(* IEC 61131-3 sources: daoli-st-library/DL_MathData (part 4) *)

(* ---- FC_DL_OrificeFlowCalc.st ---- *)
(*==============================================================================
 * 组件名称 (Component)  : FC_DL_OrificeFlowCalc
 * 所属子库 (Sublibrary) : DL_MathData
 * 当前版本 (Version)    : 1.0.0
 * 兼容性 (Platform)     : CODESYS 3.5 / TwinCAT 3 / 汇川 InoProShop / Machine Expert
 *                         仅依赖纯 IEC 61131-3 标准元素，零厂商方言
 * 功能描述 (Function)   : 孔板差压流量计算：温压补偿 + 开方 + 量程归一。
 *                         fFlow = fKCoefficient * sqrt( dP * rho(T,P) )，
 *                         密度委托 FC_DL_AirDensity（理想气体同源式，RH=0 干气口径），
 *                         开方委托 FC_DL_NthRoot(2)，本函数只做前置校验 + 钳位 + 错误码，
 *                         不重写任何开方/密度数学内核（T0 红线）。
 * 溯源 (Origin)         : 道莅 clean-room 防御性实现
 * 本文件内含 (Contains) : TYPE E_DL_MathErr / FUNCTION FC_DL_OrificeFlowCalc
 * 依赖 (Depends)        : DL_Algo/FC_DL_AirDensity、DL_MathData/FC_DL_NthRoot
 * 红线自检 (Redline)    : 无外部全局变量、无硬件地址直引 ｜ 全变量中英双语同行注释
 *                         防除零 + 量程钳位 + 非有限值防御 ｜ 枚举成员全部显式赋值
 *                         纯函数无状态保持 ｜ 输出在每条早退路径前已赋确定值
 * 错误码表 (Codes)      : 16#0001_0471 故障级 输入无效(NaN/Inf 或系数/量程非法)
 *                         16#0001_0472 故障级 差压为负
 *                         16#0001_0473 信息级 温度越界(已钳制)
 *                         16#0001_0474 信息级 压力越界(已钳制)
 *                         16#0001_0475 成功
 * 修订历史 (Revision)   : 2026-11-17  v1.0.0  首版入库 · R27 · 阶段三批 1
 * 验收向量 (Acceptance) : dP=25000 Pa, P=101325 Pa, T=20 C, K=1.0 → rho≈1.2041,
 *                         flow≈sqrt(25000*1.2041)≈173.38 m3/h，返回 0475
 *============================================================================*)

(*-----------------------------------------------------------------------------
 * 枚举: E_DL_MathErr（归属 DL_MathData，与 FC_DL_OrificeFlowCalc 同文件）
 *----------------------------------------------------------------------------*)
TYPE E_DL_MathErr :
(
    eInvalidInput := 16#0001_0471,   // 故障级：输入无效（非有限值或系数非法）/ Fault: invalid input
    eDiffPressNeg := 16#0001_0472,   // 故障级：差压为负，物理不可实现 / Fault: negative differential pressure
    eTempClamped  := 16#0001_0473,   // 信息级：温度越界已钳制 / Info: temperature clamped
    ePressClamped := 16#0001_0474,   // 信息级：压力越界已钳制 / Info: pressure clamped
    eOk           := 16#0001_0475    // 成功 / Success
);
END_TYPE

(*==============================================================================
 * 函数: FC_DL_OrificeFlowCalc（纯函数，无任何状态保持）
 * 调用约定: 每周期按需调用；返回值 = 计算有效标志。
 *============================================================================*)
FUNCTION FC_DL_OrificeFlowCalc : BOOL
VAR_INPUT
    fDiffPress_Pa  : REAL;              // 差压 [Pa]，有效域 0~50000 / Differential pressure [Pa]
    fAbsPress_Pa   : REAL;              // 绝压 [Pa]，有效域 5.0E4~2.0E6 / Absolute pressure [Pa]
    fTemp_C        : REAL;              // 温度 [摄氏度]，有效域 -40~400 / Temperature [degC]
    fKCoefficient  : REAL;              // 流量系数（含流出系数 C 的合成值），须 > 0 / Flow coefficient including discharge factor, must be > 0
    fFlowRangeMax  : REAL;              // 流量满量程 [立方米每小时]，须 > 0 / Full-scale flow [m3/h], must be > 0
END_VAR
VAR_OUTPUT
    fFlow_m3h      : REAL;              // 体积流量 [立方米每小时] / Volume flow [m3/h]
    eError         : E_DL_MathErr;      // 错误码 / Error code
END_VAR
VAR CONSTANT
    DL_ORIF_DP_MAX    : REAL := 50000.0;   // 差压量程上限 [帕] / Differential pressure span limit [Pa]
    DL_ORIF_T_MIN     : REAL := -40.0;     // 温度域下限 [摄氏度] / Temperature domain lower bound [degC]
    DL_ORIF_T_MAX     : REAL := 400.0;     // 温度域上限 [摄氏度] / Temperature domain upper bound [degC]
    DL_ORIF_P_MIN     : REAL := 5.0E4;     // 绝压域下限 [帕] / Absolute pressure lower bound [Pa]
    DL_ORIF_P_MAX     : REAL := 2.0E6;     // 绝压域上限 [帕] / Absolute pressure upper bound [Pa]
    DL_ORIF_RH_DRY    : REAL := 0.0;       // 干气口径相对湿度（委托密度入口）[%] / Dry-gas humidity fed to the density delegate [%]
    DL_ORIF_INF_MAX   : REAL := 1.0E30;    // 非有限值判定幅值上限 / Magnitude bound for finite-value check
    DL_ORIF_ZERO      : REAL := 0.0;       // 零值常量，避免裸字面量 / Zero constant, avoids a bare literal
    DL_ORIF_RHO_MIN   : LREAL := 1.0E-9;   // 密度可信下限 [千克每立方米] / Density trust lower bound [kg/m3]
END_VAR
VAR
    fDpUse    : REAL;                    // 生效差压（校验后）[帕] / Effective differential pressure [Pa]
    fTempUse  : REAL;                    // 生效温度（钳位后）[摄氏度] / Effective temperature [degC]
    fPressUse : REAL;                    // 生效绝压（钳位后）[帕] / Effective absolute pressure [Pa]
    fRho      : LREAL;                   // 委托密度输出 [千克每立方米] / Density from the delegate [kg/m3]
    fRadicand : LREAL;                   // 开方被开方数 [帕·千克每立方米] / Radicand [Pa*kg/m3]
    fRootVal  : LREAL;                   // 委托开方输出 [无量纲合成] / Square root from the delegate
    bRootOk   : BOOL;                    // 委托开方有效标志 / Delegate root validity flag
    bNonFin   : BOOL;                    // 非有限输入汇总标志 / Non-finite input aggregate flag
END_VAR

(*------------------------------------------------------------------------------
 * 段 1｜出口默认值：任何早退路径前输出已确定（哨兵 0 流量 + 输入无效码）
 *----------------------------------------------------------------------------*)
FC_DL_OrificeFlowCalc := FALSE;                       // 返回值默认无效 / return defaults to invalid
fFlow_m3h := DL_ORIF_ZERO;                            // 流量哨兵 0 / flow sentinel zero
eError := E_DL_MathErr.eInvalidInput;                 // 默认输入无效码 / default invalid-input code

(*------------------------------------------------------------------------------
 * 段 2｜非有限值闸：NaN 用自反判（x <> x），溢出用幅值上限判
 *----------------------------------------------------------------------------*)
bNonFin := (fDiffPress_Pa <> fDiffPress_Pa) OR (ABS(fDiffPress_Pa) > DL_ORIF_INF_MAX)
        OR (fAbsPress_Pa  <> fAbsPress_Pa)  OR (ABS(fAbsPress_Pa)  > DL_ORIF_INF_MAX)
        OR (fTemp_C       <> fTemp_C)       OR (ABS(fTemp_C)       > DL_ORIF_INF_MAX)
        OR (fKCoefficient <> fKCoefficient) OR (ABS(fKCoefficient) > DL_ORIF_INF_MAX)
        OR (fFlowRangeMax <> fFlowRangeMax) OR (ABS(fFlowRangeMax) > DL_ORIF_INF_MAX);
IF bNonFin THEN
    RETURN;                                           // 早退：保持默认输出 / early exit with defaults
END_IF

(*------------------------------------------------------------------------------
 * 段 3｜配置与符号闸：系数/量程必须为正，差压不允许为负
 *----------------------------------------------------------------------------*)
IF (fKCoefficient <= DL_ORIF_ZERO) OR (fFlowRangeMax <= DL_ORIF_ZERO) THEN
    RETURN;                                           // 配置非法：保持输入无效码 / invalid configuration
END_IF
IF fDiffPress_Pa < DL_ORIF_ZERO THEN
    eError := E_DL_MathErr.eDiffPressNeg;             // 故障级：差压为负 / fault: negative dp
    RETURN;
END_IF
fDpUse := fDiffPress_Pa;                              // 差压非负直接采用 / non-negative dp adopted

(*------------------------------------------------------------------------------
 * 段 4｜温度/压力钳位（信息级越界码，先到先得但压力优先级低：温度先判）
 *----------------------------------------------------------------------------*)
eError := E_DL_MathErr.eOk;                           // 预置成功 / preset success
fTempUse := fTemp_C;                                  // 温度工作副本 / temperature working copy
IF fTempUse < DL_ORIF_T_MIN THEN
    fTempUse := DL_ORIF_T_MIN;                        // 下限钳位 / floored
    eError := E_DL_MathErr.eTempClamped;              // 信息级：温度越界 / info: temperature clamped
ELSIF fTempUse > DL_ORIF_T_MAX THEN
    fTempUse := DL_ORIF_T_MAX;                        // 上限钳位 / capped
    eError := E_DL_MathErr.eTempClamped;              // 信息级：温度越界 / info: temperature clamped
END_IF
fPressUse := fAbsPress_Pa;                            // 压力工作副本 / pressure working copy
IF fPressUse < DL_ORIF_P_MIN THEN
    fPressUse := DL_ORIF_P_MIN;                       // 下限钳位 / floored
    IF eError = E_DL_MathErr.eOk THEN
        eError := E_DL_MathErr.ePressClamped;         // 信息级：压力越界（不覆盖温度码）/ info: pressure clamped
    END_IF
ELSIF fPressUse > DL_ORIF_P_MAX THEN
    fPressUse := DL_ORIF_P_MAX;                       // 上限钳位 / capped
    IF eError = E_DL_MathErr.eOk THEN
        eError := E_DL_MathErr.ePressClamped;         // 信息级：压力越界（不覆盖温度码）/ info: pressure clamped
    END_IF
END_IF

(*------------------------------------------------------------------------------
 * 段 5｜委托密度（理想气体同源式，RH=0 干气口径；委托 FC_DL_AirDensity）
 *----------------------------------------------------------------------------*)
fRho := FC_DL_AirDensity(fTempC := REAL_TO_LREAL(fTempUse), fPressPa := REAL_TO_LREAL(fPressUse), fRh := REAL_TO_LREAL(DL_ORIF_RH_DRY));   // 密度委托 [千克每立方米] / density via delegate
IF (fRho <> fRho) OR (ABS(fRho) > REAL_TO_LREAL(DL_ORIF_INF_MAX)) OR (fRho <= DL_ORIF_RHO_MIN) THEN
    eError := E_DL_MathErr.eInvalidInput;             // 委托输出不可信：按输入无效处置 / unusable delegate output
    fFlow_m3h := DL_ORIF_ZERO;                        // 流量哨兵 / flow sentinel
    FC_DL_OrificeFlowCalc := FALSE;                   // 返回无效 / return invalid
    RETURN;
END_IF

(*------------------------------------------------------------------------------
 * 段 6｜委托开方（FC_DL_NthRoot(2)）：被开方数 = 差压 x 密度，段 5 已保证非负
 *----------------------------------------------------------------------------*)
fRadicand := REAL_TO_LREAL(fDpUse) * fRho;                     // 被开方数 [帕·千克每立方米] / radicand
fRootVal := FC_DL_NthRoot(fValue := fRadicand, nRoot := 2, bValid => bRootOk);   // 开方委托 / root via delegate
IF (NOT bRootOk) OR (fRootVal <> fRootVal) OR (ABS(fRootVal) > REAL_TO_LREAL(DL_ORIF_INF_MAX)) THEN
    eError := E_DL_MathErr.eInvalidInput;             // 委托失败按输入无效处置 / delegate failure mapped to invalid input
    FC_DL_OrificeFlowCalc := FALSE;                   // 返回无效 / return invalid
    RETURN;
END_IF

(*------------------------------------------------------------------------------
 * 段 7｜量程换算与上限钳制：flow = K x root，超出满量程钳制并保留成功码
 *----------------------------------------------------------------------------*)
fFlow_m3h := LREAL_TO_REAL(fRootVal) * fKCoefficient;   // 合成流量 [立方米每小时] / composed flow [m3/h]
IF fFlow_m3h > fFlowRangeMax THEN
    fFlow_m3h := fFlowRangeMax;                       // 满量程钳制 / clamped to full scale
END_IF
IF fFlow_m3h < DL_ORIF_ZERO THEN
    fFlow_m3h := DL_ORIF_ZERO;                        // 下限防护（禁止伪负流量）/ floor guard
END_IF
FC_DL_OrificeFlowCalc := TRUE;                        // 计算有效 / computation valid
RETURN;
END_FUNCTION

(* ---- FC_DL_ParityCalc.st ---- *)
(*
    FC_DL_ParityCalc —— 奇/偶校验位计算（位宽显式参数 + 无效位宽拒算）
    ------------------------------------------------------------------
    分类      : DL_MathData / Data-Integrity
    前缀      : FC_DL_
    版本      : 1.0.0
    来源标签  : iec-std-wrapper（T0）
    溯源      : IEC 61131-3 标准语义的道莅防御性实现
                （纯位运算循环，无内建校验内核依赖；未复制任何闭源厂商源码）
    平台      : 纯 IEC 61131-3，CODESYS / TwinCAT / InoProShop 通用
    分工声明  : 与存量 FC_DL_LwordBitCount（位计数）、FC_DL_Crc16Generic（CRC 族）
                分工——BitCount 返回置位总数，本件只做奇/偶校验位单出口；
                CRC 为多项式校验，与本件奇偶口径互不替代。
    作者      : 道莅代码库 · PLC 编程专家（R57）
    ------------------------------------------------------------------
    功能说明  : 对 LWORD 数据低 nWidth 位计算奇/偶校验位。位宽域 [1, 64]，
                越域拒算置错误（等效钳位语义：非法值不执行任何位运算）；
                偶校验 = 置位总数模 2；奇校验 = 偶校验取反。移位量恒为 1，
                结构性安全（R48）。
    错误码    : 0000 正常 / 16#0003_0005 位宽越域拒算
    修订记录  : 2026-11-21 v1.0.0 首次入库（R57 批 3 · 序号 13）
*)
TYPE E_DL_ParityMode :
(
    eEven := 0, // 偶校验：置位总数为偶时校验位 0 / even parity, a zero bit when the set count is even
    eOdd  := 1  // 奇校验：置位总数为奇时校验位 0 / odd parity, a zero bit when the set count is odd
);
END_TYPE

FUNCTION FC_DL_ParityCalc : BOOL
VAR_INPUT
    uData  : LWORD; // 被校验数据（仅低 nWidth 位参与）[-] / the checked data, only the low nWidth bits participate
    nWidth : INT;   // 参与校验的位宽 [位]，域 1..64 / the participating width [bit], one through sixty four
    eMode  : E_DL_ParityMode := E_DL_ParityMode.eEven; // 校验模式 [枚举] / the parity mode [enum]
END_VAR
VAR_OUTPUT
    eErr   : UDINT; // 错误码，0 = 正常 / error code, zero is ok
    bError : BOOL;  // 出错标志，eErr 非 0 时为真 / error flag, true when eErr is nonzero
    bValid : BOOL;  // 结果是否可用，拒算时为假 / the result usable, false when rejected
END_VAR
VAR
    uMask  : LWORD; // 位测试掩码 [-] / the bit test mask
    nI     : INT;   // 循环计数 [位] / the loop counter
    nOnes  : INT;   // 置位总数 [个] / the set bit count
    bBit   : BOOL;  // 当前位为 1 [-] / the current bit set
END_VAR

// 段 1｜返回值与错误状态预置安全值（四段式第一段，R45）/ segment 1, preset the return and error states
FC_DL_ParityCalc := FALSE; // 校验位预置 0 / preset the parity bit to zero
eErr   := 16#0000_0000; // 错误码预置正常 / preset the code to ok
bError := FALSE; // 错误标志预置假 / preset the error flag false
bValid := TRUE; // 有效标志预置真 / preset the valid flag true

// 段 2｜位宽域闸：越域拒算（边界十三）/ segment 2, the width gate, out of domain rejects
IF (nWidth < 1) OR (nWidth > 64) THEN // 位宽非法 / an illegal width
    eErr   := 16#0003_0005; // 错误级：位宽越域拒算 / error grade, an out of domain width rejected
    bError := TRUE; // 置错误标志 / raise the error flag
    bValid := FALSE; // 输出不可用 / the output void
    RETURN; // 返回预置安全值 FALSE / return the preset safe false
END_IF

// 段 3｜逐位测试计数：移位量恒 1，结构性安全（R48）/ segment 3, the bit by bit tally, the shift amount always one
uMask := LWORD#1; // 掩码从最低位起步 / the mask starts at the lowest bit
nOnes := 0; // 置位计数清零 / clear the tally
FOR nI := 1 TO nWidth DO // 有界循环（nWidth 已证 1..64）/ the bounded loop
    bBit := (uData AND uMask) <> LWORD#0; // 当前位测试 / the current bit test
    IF bBit THEN // 置位 / a set bit
        nOnes := nOnes + 1; // 计数推进 / advance the tally
    END_IF
    IF nI < nWidth THEN // 末位后不再移位（防 64 位移出丢失语义位）/ no shift after the last bit
        uMask := SHL(uMask, 1); // 掩码左移 1 位（移位量常量）/ shift the mask left by one
    END_IF
END_FOR

// 段 4｜奇偶模式判定（nOnes 非负，MOD 合法）/ segment 4, the parity verdict, the modulus on a nonnegative tally
IF eMode = E_DL_ParityMode.eEven THEN // 偶校验 / the even mode
    FC_DL_ParityCalc := (nOnes MOD 2) = 1; // 置位总数为奇时校验位 1 / the parity bit one on an odd tally
ELSIF eMode = E_DL_ParityMode.eOdd THEN // 奇校验 / the odd mode
    FC_DL_ParityCalc := (nOnes MOD 2) = 0; // 置位总数为偶时校验位 1 / the parity bit one on an even tally
ELSE // 非法模式兜底 / the illegal mode fallback
    eErr   := 16#0003_0005; // 错误级：模式非法拒算 / error grade, an illegal mode rejected
    bError := TRUE; // 置错误标志 / raise the error flag
    bValid := FALSE; // 输出不可用 / the output void
    FC_DL_ParityCalc := FALSE; // 返回安全值 / return the safe value
END_IF
END_FUNCTION

(* ---- FC_DL_PercentileRank.st ---- *)
(*
  ==================================================================
  组件名 Component  : FC_DL_PercentileRank
  分类   Category   : DL_MathData
  前缀   Naming     : FC_DL_ ｜ b/n/u/f/t/e/st 类型前缀制（R265）
  码位   Code ID    : 16#0001_0653（信息级）｜ 16#0001_0654 / 0656（故障级）
  版本   Version    : 1.0.1
  复杂度 Complexity  : 中
  功能   Purpose    : 值 → 百分位排名（0..100），即「当前值在历史分布中的位置」，
                      SPC / 过程能力定位用；三口径（弱 / 强 / 中位排名）显式可选。
  开源溯源 Origin    : IEC 61131-3 标准语义的道莅防御性实现（clean-room，无第三方代码行）
  许可证 License    : MIT
  参考   Reference  : IEC 61131-3:2013 §6.6 标准运算符与 §6.6.1 比较/选择语义
  平台   Platform   : 纯 IEC 61131-3（FOR / CASE / 四则 / 委托），三平台通用
  依赖   Depends    : FC_DL_SortIndexLReal（索引排序属主，本件委托排序，R140）
  分工声明 Split     : FC_DL_PercentileLReal（分位→值）/ FC_DL_WeightedPercentile（加权分位）
                      / FC_DL_QuantileCalc（分位族通用）为「分位 → 值」方向；本件是逆运算
                      「值 → 分位」。选型差异：限值设定用分位→值（给定分位求门限值），
                      SPC 定位用本件（给定实测值求它落在历史分布的哪一档）（R216 双向互引）。
  归属 Ownership     : E_DL_RankMethod 属主为本文件（全库唯一定义，R264）；引用件只引用
                      不重声明。委托件码位随其属主回传（R66）。
  ------------------------------------------------------------------
  边界 Boundary     :
                      一 有效样本口径：非有限（NaN / ±Inf）样本逐条剔除并计入局部 nNonFinite，
                         全部判据的除子一律用剔除后的 nEff，禁用 nCount 直接作除子；
                         nNonFinite 口径定稿（v1.0.1 返修 R63 · 修 R62-D7 轻）：**不外显**
                         （维持局部留档、不出现在输出契约），剔除诊断请用
                         FC_DL_SignalStatistics（非有限样本计数口径属主）；
                      二 nCount 越域（< 1 或 > 256）判故障早退；剔除后 nEff = 0 同码处置
                         （两场景在出口上同为「无可排名样本」，合并为一码，R90 反证句见码表）；
                      三 fValue 非有限（NaN / ±Inf）判故障早退，禁把 NaN 当合格值参与比较；
                      四 排名口径非法（枚举越域）由 CASE ... ELSE 拦为 eMidRank 并置信息级
                         组态码，禁静默；
                      五 三口径公式：eWeak = nBelow / nEff；eStrong = (nBelow + nEqual) / nEff；
                         eMidRank = (nBelow + nEqual / 2) / nEff；全乘 100 得 [%]；
                      六 浮点判等只用于「与待定位值相等」的容差判定，禁用 = / <> 判等；
                      七 委托返回值与 bValid 由两个独立变量承接后合取（R62-D5 教训）；
                      八 纯函数：无记忆量、无定时器、无边沿实例，每调用重算。
  错误码 Codes      :
    16#0001_0653【信息级】排名口径枚举越域，已落中位排名口径（不置 bError）
    16#0001_0654【故障级】有效样本数越域：nCount < 1 或 > 256，或剔除非有限后 nEff = 0
    16#0001_0656【故障级】数值非有限：fValue 为 NaN / ±Inf，或结果复检命中非有限（后者理论上不可达的兜底分支）
  码位反证 Note     :
    0654 合并「入参越域」与「剔净后为空」的理由：两者的出口组合完全相同（均为
    nBelow = 0、nEqual = 0、fPct = 0、bValid = FALSE），三组以内输出无法唯一还原该场景，
    按 R90 不另立码；0656 不可并入 0654，因 bValid 与 nEff 在两种场景下可唯一区分
    （前者 nEff ≥ 1、后者 nEff = 0）；0656 同时承担结果复检兜底：该分支与「fValue 非有限」
    在出口上完全同形（fPct = 0、bValid = FALSE、nBelow / nEqual 保持计数），三组以内输出
    无法区分，故按 R90 共用一码而不另立。
  验收 Acceptance   :
    算法已证（脚本）：未跑 ｜ 编译器已证（三平台）：未跑
    V1 全同样本、fValue 相等 → eWeak 0 / eStrong 100 / eMidRank 50（逐口径断言）
    V2 fValue 小于最小样本 → 0%；V3 大于最大样本 → 100%
    V4 单样本 nCount = 1 → 三口径 0 / 100 / 50
    V5 含 2 个 NaN + 6 个有效 → nEff = 6（除子已证 ≥ 1），排名按 6 计
    V6 nCount = 0 → 码 0654 + 早退（禁除零）；V7 nCount = 257 → 同码早退
    V8 eMethod = 99（非法枚举）→ 落 eMidRank + 码 0653（bError = FALSE）
    V9 fValue = NaN → 码 0656 + bValid = FALSE
  修订记录 Revision  :
    2026-11-21  v1.0.0  R62 首版（批 3 · 序号 8）
    2026-11-21  v1.0.1  R63 返修 R5（R62-D7 轻）：nNonFinite 口径二选一定稿为「不外显」，
                        头注释与声明行注明诊断请用 FC_DL_SignalStatistics（不改接口）
  ==================================================================
*)
TYPE E_DL_RankMethod :
(
    eWeak    := 0, // 弱排名：只计严格小于的样本（同值全落上沿，保守低估）/ the weak rank counting strictly smaller samples only
    eStrong  := 1, // 强排名：计小于与相等的样本（同值全落上沿，偏乐观）/ the strong rank counting smaller and equal samples
    eMidRank := 2  // 中位排名：相等样本各计一半（同值取中点，统计口径最中性）/ the mid rank giving half credit to equal samples
);
END_TYPE

FUNCTION FC_DL_PercentileRank : BOOL
VAR_IN_OUT
    afSamples : ARRAY[0..255] OF LREAL; // 样本序列 [工程单位]，只读 / the sample series, read only
END_VAR
VAR_INPUT
    nCount  : DINT := 0;                          // 有效样本数入参 [个]，合法域 1..256 / the sample count, legal one to two hundred fifty six
    fValue  : LREAL := 0.0;                       // 待定位值 [工程单位]，必须有限 / the value to locate, must be finite
    eMethod : E_DL_RankMethod := E_DL_RankMethod.eMidRank; // 排名口径 [-] / the ranking convention
END_VAR
VAR_OUTPUT
    fPct   : LREAL; // 百分位排名 [%]，0..100 / the percentile rank in percent
    nBelow : DINT;  // 严格小于待定位值的样本数 [个] / the count of samples strictly below the value
    nEqual : DINT;  // 与待定位值相等的样本数 [个] / the count of samples equal to the value
    bValid : BOOL;  // 结果可用 [-] / the result usable flag
    eErr   : UDINT; // 错误码，0 = 正常 / the error code, zero is ok
    bError : BOOL;  // 错误标志，故障级码置位（R45 配对）/ the error flag raised with a fault level code
END_VAR
VAR
    aVal      : ARRAY[0..255] OF LREAL;        // 剔除非有限后的有效样本副本 [工程单位] / the finite sample copy
    aIdx      : ARRAY[0..255] OF DINT;         // 委托输出的排序索引排列 [下标] / the sorted permutation from the delegate
    k         : DINT := 0;                     // 遍历索引 [下标] / the traversal index
    nEff      : DINT := 0;                     // 剔除非有限后的有效样本数 [个]（除子）/ the effective sample count used as the divisor
    nNonFinite: DINT := 0;                     // 剔除的非有限样本数 [个]（仅局部留档，不外显不作除子，v1.0.1 定稿；诊断请用 FC_DL_SignalStatistics）/ the dropped non finite sample count, local only and never exposed, use the signal statistics component for diagnostics
    nCountUse : DINT := 0;                     // 钳位前的入参样本数接管量 [个] / the raw input count before the domain gate
    fPctUse   : LREAL := 0.0;                  // 排名百分比工作副本 [%] / the working percentile copy
    eUse      : E_DL_RankMethod := E_DL_RankMethod.eMidRank; // 归一后的排名口径 [-] / the normalized ranking convention
    bSortRet  : BOOL := FALSE;                 // 委托返回值承接量（独立承接）/ the delegate return holder
    bSortValid: BOOL := FALSE;                 // 委托 bValid 承接量（独立承接）/ the delegate valid holder
    uSortErr  : UDINT := 16#0000_0000;         // 委托错误码承接量 [码] / the delegate error code holder
    bSortErr  : BOOL := FALSE;                 // 委托故障位承接量 / the delegate fault bit holder
    bSortOk   : BOOL := FALSE;                 // 返回值与可用位合取后的排序可用位 / the conjunction of the return value and the valid flag
END_VAR  // R64 结构补齐：VAR 段缺失的 END_VAR（门禁机械修复）
VAR CONSTANT
    DL_PRK_NMAX : DINT := 256;         // 样本容量上界 [个]，与数组容量一致 / the capacity aligned with the array
    DL_PRK_ONE : DINT := 1;            // 整型一常量 [个] / the integer one constant
    DL_PRK_ZERO : DINT := 0;           // 整型零常量 [个] / the integer zero constant
    DL_PRK_PCT100 : LREAL := 100.0;    // 百分制换算系数 [%] / the percent scaling factor
    DL_PRK_HALF : LREAL := 2.0;        // 相等样本折半除子 [-] / the halving divisor for the equal samples
    DL_PRK_EQEPS : LREAL := 1.0E-6;    // 相等判定容差 [工程单位]，禁用 = / <> 判等 / the equality tolerance, plain equality operators are forbidden
END_VAR

// 段 1｜返回值与全部出口预置安全值（R45 四段式第一段）+ 局部量显式预置（R254）/ segment 1, the preset
FC_DL_PercentileRank := FALSE; // 返回值预置假 / preset the return false
fPct := 0.0; // 百分比预置零 [%] / preset the percentage zero
nBelow := 0; // 小于计数预置零 [个] / preset the below count zero
nEqual := 0; // 相等计数预置零 [个] / preset the equal count zero
bValid := FALSE; // 可用标志预置假 / preset the validity false
eErr := 16#0000_0000; // 错误码预置正常 / preset the code to ok
bError := FALSE; // 错误标志预置假 / preset the error flag false
nEff := DL_PRK_ZERO; // 有效样本数预置零 [个] / preset the effective count zero
nNonFinite := DL_PRK_ZERO; // 剔除计数预置零 [个] / preset the dropped count zero
nCountUse := DL_PRK_ZERO; // 入参计数接管量预置零 [个] / preset the raw count holder zero
fPctUse := 0.0; // 百分比工作副本预置零 [%] / preset the working copy zero
bSortRet := FALSE; // 委托返回值承接量预置假 / preset the return holder false
bSortValid := FALSE; // 委托可用位承接量预置假 / preset the valid holder false
uSortErr := 16#0000_0000; // 委托码承接量预置零 [码] / preset the delegate code zero
bSortErr := FALSE; // 委托故障位承接量预置假 / preset the delegate fault holder false
bSortOk := FALSE; // 排序可用位预置假 / preset the sort usable bit false
eUse := E_DL_RankMethod.eMidRank; // 口径工作量预置中位排名（偏保守的中性口径）/ preset the convention to the neutral mid rank

// 段 2｜样本数域闸（边界二，早退禁除零）/ segment 2, the sample count domain gate
nCountUse := nCount; // 入参计数接管 [个] / take the raw count
IF (nCountUse < DL_PRK_ONE) OR (nCountUse > DL_PRK_NMAX) THEN // 计数越域 / the count is out of the domain
    eErr := 16#0001_0654; // 故障级：有效样本数越域 / fault grade, the effective sample count is out of the domain
    bError := TRUE; // 同拍置故障标志（R45 配对）/ raise the fault flag on the same scan
    bValid := FALSE; // 结果不可用 / the result is not usable
    RETURN; // 早退，绝不进入除法 / early return, no division is ever reached
END_IF

// 段 3｜待定位值非有限闸（边界三，NaN 与 ±Inf 逐个点名，R272）/ segment 3, the value finiteness gate
IF (fValue <> fValue) OR ((fValue - fValue) <> (fValue - fValue)) THEN // NaN 或 ±Inf / NaN or an infinity
    eErr := 16#0001_0656; // 故障级：待定位值非有限 / fault grade, the value to locate is not finite
    bError := TRUE; // 同拍置故障标志（R45 配对）/ raise the fault flag on the same scan
    bValid := FALSE; // 结果不可用 / the result is not usable
    RETURN; // 早退 / early return
END_IF

// 段 4｜样本非有限剔除（边界一：除子口径 = 有效样本数，绝不用入参计数作除子）/ segment 4, drop the non finite samples
FOR k := 0 TO nCountUse - 1 DO // 有界遍历（上界已证 ≤ 256）/ the bounded traversal with a proven ceiling
    IF (afSamples[k] = afSamples[k]) AND ((afSamples[k] - afSamples[k]) = (afSamples[k] - afSamples[k])) THEN // 有限样本 / a finite sample
        aVal[nEff] := afSamples[k]; // 有限样本写入副本 [工程单位] / copy the finite sample
        nEff := nEff + DL_PRK_ONE; // 有效计数推进 [个] / advance the effective count
    ELSE // 非有限样本 / a non finite sample
        nNonFinite := nNonFinite + DL_PRK_ONE; // 剔除计数推进 [个] / advance the dropped count
    END_IF
END_FOR
IF nEff < DL_PRK_ONE THEN // 剔净后无可排名样本（与段 2 同码，出口组合不可区分，R90）/ no sample remains after the drop
    eErr := 16#0001_0654; // 故障级：有效样本数越域（此处为剔净后为空）/ fault grade, the effective count is empty after the drop
    bError := TRUE; // 同拍置故障标志（R45 配对）/ raise the fault flag on the same scan
    bValid := FALSE; // 结果不可用 / the result is not usable
    RETURN; // 早退，除子已证 ≥ 1 才允许进入段 6 / early return, the divisor is proven at least one before the percentage segment
END_IF

// 段 5｜委托索引排序（R140；返回值与可用位分承后合取，R62-D5）/ segment 5, the delegated index sort
bSortRet := FC_DL_SortIndexLReal(afValues := aVal, nCount := nEff, aIdx => aIdx, bValid => bSortValid, eErr => uSortErr, bError => bSortErr); // 委托排序：两路各自承接 / delegate the sort into two distinct holders
bSortOk := bSortRet AND bSortValid; // 返回值与可用位合取（IEC 未规定两者的求值次序）/ conjoin the two signals since their evaluation order is unspecified
IF (NOT bSortOk) OR bSortErr THEN // 委托失败 / the delegate failed
    eErr := uSortErr; // 委托码回传（码随属主，R66）/ replay the delegate code
    bError := bSortErr; // 委托故障位回传 / replay the delegate fault bit
    bValid := FALSE; // 结果不可用 / the result is not usable
    RETURN; // 早退 / early return
END_IF

// 段 6｜排名计数（小于 / 相等，相等用容差判定，禁判等算符）/ segment 6, the rank counting with a tolerance equality test
FOR k := 0 TO nEff - 1 DO // 按排序序有界遍历 / the bounded traversal in the sorted order
    IF aVal[aIdx[k]] < fValue THEN // 严格小于 / strictly below
        nBelow := nBelow + DL_PRK_ONE; // 小于计数推进 [个] / advance the below count
    ELSIF ABS(aVal[aIdx[k]] - fValue) < DL_PRK_EQEPS THEN // 容差相等（浮点禁判等）/ equality inside the tolerance
        nEqual := nEqual + DL_PRK_ONE; // 相等计数推进 [个] / advance the equal count
    END_IF
END_FOR

// 段 7｜排名口径归一并计算百分比（边界四，CASE 必带 ELSE 兜底）/ segment 7, the convention normalization and the percentage
CASE eMethod OF
    E_DL_RankMethod.eWeak: // 弱排名口径 / the weak rank convention
        eUse := E_DL_RankMethod.eWeak; // 口径接管 / take the convention
        fPctUse := (DINT_TO_LREAL(nBelow) / DINT_TO_LREAL(nEff)) * DL_PRK_PCT100; // 弱排名百分比 [%] / the weak rank percentage
    E_DL_RankMethod.eStrong: // 强排名口径 / the strong rank convention
        eUse := E_DL_RankMethod.eStrong; // 口径接管 / take the convention
        fPctUse := ((DINT_TO_LREAL(nBelow) + DINT_TO_LREAL(nEqual)) / DINT_TO_LREAL(nEff)) * DL_PRK_PCT100; // 强排名百分比 [%] / the strong rank percentage
    E_DL_RankMethod.eMidRank: // 中位排名口径 / the mid rank convention
        eUse := E_DL_RankMethod.eMidRank; // 口径接管 / take the convention
        fPctUse := ((DINT_TO_LREAL(nBelow) + (DINT_TO_LREAL(nEqual) / DL_PRK_HALF)) / DINT_TO_LREAL(nEff)) * DL_PRK_PCT100; // 中位排名百分比 [%] / the mid rank percentage
    ELSE // 非法枚举值：落中位排名并置组态码（禁静默，边界四）/ an illegal enumeration falls back to the mid rank with a code
        eUse := E_DL_RankMethod.eMidRank; // 落中性口径 / fall back to the neutral convention
        fPctUse := ((DINT_TO_LREAL(nBelow) + (DINT_TO_LREAL(nEqual) / DL_PRK_HALF)) / DINT_TO_LREAL(nEff)) * DL_PRK_PCT100; // 中位排名百分比 [%] / the mid rank percentage
        eErr := 16#0001_0653; // 信息级：排名口径越域，已落中位排名 / informational, the convention is out of the domain and the mid rank was used
        bError := FALSE; // 信息级不置故障标志（R285）/ keep the error flag false, this is informational
END_CASE

// 段 8｜结果复检兜底（结果非有限必三件套，R258）/ segment 8, the result recheck with the three part fallback
IF (fPctUse <> fPctUse) OR ((fPctUse - fPctUse) <> (fPctUse - fPctUse)) THEN // 结果非有限（理论上不可达，防御保留）/ a non finite result, unreachable by theory, kept as a defence
    fPct := 0.0; // 兜底安全值 [%] / the bottom line safe value
    eErr := 16#0001_0656; // 故障级：待定位值非有限（同族三件套口径）/ fault grade under the same family code
    bError := TRUE; // 置故障标志（R45 配对）/ raise the fault flag
    bValid := FALSE; // 结果不可用 / the result is not usable
    RETURN; // 早退 / early return
END_IF

// 段 9｜统一出口 / segment 9, the unified outlet
fPct := fPctUse; // 百分比出口 [%] / the percentage outlet
bValid := TRUE; // 结果可用 / the result is usable
FC_DL_PercentileRank := TRUE; // 返回成功 / return success
END_FUNCTION

(* ---- FC_DL_PolarTransform2D.st ---- *)
(*==============================================================================
 * 组件名称 (Component)  : FC_DL_PolarTransform2D
 * 所属子库 (Sublibrary) : DL_MathData
 * 前缀     (Prefix)     : FC_DL_
 * 当前版本 (Version)    : 1.0.0
 * 兼容性   (Platform)   : CODESYS 3.5 / TwinCAT 3 / 汇川 InoProShop / Schneider
 *                         Machine Expert；纯 IEC 61131-3（第 3 版），
 *                         仅依赖标准函数 SQRT / ATAN2 / COS / SIN / ABS / TRUNC，
 *                         零厂商方言、无状态纯函数
 * 作者     (Author)     : 道莅代码库 · PLC编程专家（R31）
 * 开源溯源 (Origin)     : 直角坐标与极坐标双向变换公开数学语义，
 *                         IEC 61131-3 标准语义的道莅防御性实现，
 *                         防平方溢出归一范式借鉴本库 CalcDistance3D 行为定义，
 *                         未复制任何外部源码行
 * 功能描述 (Function)   : 直角坐标与极坐标双向变换纯函数。正变换输出半径与
 *                         角度（角度单位 deg，值域 0..360）；先取最大分量归一
 *                         防平方溢出；逆变换先做角度归一防大角度精度损失。
 *                         原点正变换合法（r=0、theta=0 写死本头注释）；负半径
 *                         语义歧义按非法拒绝，不替调用方裁定方向。
 * 码位     (Codes)      : 16#0001_0092 信息级：输入非有限（不置故障标志）
 *                         16#0001_0093 信息级：负半径非法拒绝
 *                         16#0001_0094 信息级：角度超域已归一钳位
 *                         16#0001_0095 信息级：变换模式非法（ELSE 兜底拒绝）
 *                         纯函数四槽全信息级：拒绝时 bValid=FALSE 表达不可用，
 *                         不设故障标志引脚（规格 §2 裁定，FC 无故障级语义）。
 * 边界防错 (Boundary)   : 1 非有限判据：x<>x 自反判 NaN 加幅值界双侧判 Inf；
 *                         2 正变换 m=MAX(ABS(x),ABS(y)) 归一后再求平方和；
 *                         3 ATAN2(0,0) 无定义，原点单列直取 theta=0；
 *                         4 角度一律换算为 deg 并归一到 0..360 半开区间；
 *                         5 大角度先取模归一，防三角函数精度损失。
 * 修订历史 (Revision)   : 2026-11-18 v1.0.0 首版入库（R31 · 阶段三 · 序 2）
 *==============================================================================*)

(*------------------------------------------------------------------------------
 * 枚举: E_DL_PolarMode（归属本函数，同文件发布，全库唯一属主）
 *----------------------------------------------------------------------------*)
TYPE E_DL_PolarMode :
(
    eToPolar := 0,    // 正变换：直角转极，输出半径/角度 deg / To polar, radius and angle in deg
    eToCart  := 1     // 逆变换：极转直角，输入半径/角度 deg / To cartesian, radius and angle in deg
);
END_TYPE

(*==============================================================================
 * 函数: FC_DL_PolarTransform2D（纯函数，无状态，同输入必得同输出）
 *==============================================================================*)
FUNCTION FC_DL_PolarTransform2D : BOOL
VAR_INPUT
    fX      : LREAL;                    // 直角模式：X 坐标；极模式：半径 [mm 或调用方单位] / Cartesian X or radius
    fY      : LREAL;                    // 直角模式：Y 坐标；极模式：角度 [deg] / Cartesian Y or angle in deg
    eMode   : E_DL_PolarMode;           // 变换方向选择 / Transformation direction selector
END_VAR
VAR_OUTPUT
    fA      : LREAL;                    // 极模式输出：半径；直角模式输出：X [同输入单位] / Radius or X output
    fB      : LREAL;                    // 极模式输出：角度 [deg]；直角模式输出：Y [同输入单位] / Angle deg or Y output
    bValid  : BOOL;                     // 结果可用标志 / Result validity flag
    uErrorId : UINT;                    // 信息级码，0 = 无信息 / Info code, 0 = none
END_VAR
VAR
    fMaxC   : LREAL;                    // 最大分量模，防平方溢出归一基准 / Max component magnitude
    fXn     : LREAL;                    // 归一后 X 分量 / Normalised X component
    fYn     : LREAL;                    // 归一后 Y 分量 / Normalised Y component
    fRad    : LREAL;                    // 中间角 [rad] / Intermediate angle [rad]
    fDeg    : LREAL;                    // 中间角 [deg]，归一前 / Intermediate angle [deg] before normalising
    fLim    : LREAL;                    // 有限幅值判界复用寄存 / Finiteness bound register
END_VAR
VAR CONSTANT
    DL_POL_PI     : LREAL := 3.14159265358979323846; // 圆周率 / Pi constant
    DL_POL_DEG180 : LREAL := 180.0;                  // 弧度转角度系数 [deg/rad] / Rad to deg factor
    DL_POL_EPS    : LREAL := 1.0E-300;               // 原点判零容差 / Origin zero tolerance
    DL_POL_FIN    : LREAL := 1.7976931348623157E308; // LREAL 幅值上限 / LREAL magnitude ceiling
    DL_POL_ANGMAX : LREAL := 1.0E6;                  // 角度超域判界 [deg]，超界先取模 / Angle range bound [deg] before modulo
END_VAR

// ---- 段 1｜出口默认值：入口即赋确定值，提前 RETURN 前输出已确定 ---------------
FC_DL_PolarTransform2D := TRUE;                       // 返回值默认真，拒绝时显式改 FALSE / Preset TRUE, set FALSE on rejection
fA      := 0.0;                                       // 输出 A 预置零 / Preset output A
fB      := 0.0;                                       // 输出 B 预置零 / Preset output B
bValid  := FALSE;                                     // 可用标志预置假 / Preset invalid
uErrorId := 16#0000;                                  // 信息码清零（UINT 16 位段）/ Clear info code
fLim    := DL_POL_FIN;                                // 判界装载 / Load finiteness bound

// ---- 段 2｜非有限防御：NaN 用 x<>x 自反判，Inf 用幅值双侧判 -------------------
IF (fX <> fX) OR (fY <> fY) OR (ABS(fX) >= fLim) OR (ABS(fY) >= fLim) THEN
    uErrorId := 16#0001_0092;                         // 信息级：输入非有限 / Info: non-finite input
    RETURN;                                           // 拒绝出口，输出保持预置零 / Rejection exit with deterministic zeros
END_IF

// ---- 段 3｜按模式分派（CASE 含 ELSE 非法模式兜底）---------------------------
CASE eMode OF
    eToPolar:
        // 正变换：先取最大分量归一，防 x^2+y^2 溢出（CalcDistance3D 范式）
        fMaxC := MAX(ABS(fX), ABS(fY));               // 最大分量模 / Max component magnitude
        IF fMaxC < DL_POL_EPS THEN
            fA := 0.0;                                // 原点正变换合法：r=0 写死头注释 / Origin is legal, r=0
            fB := 0.0;                                // 原点正变换合法：theta=0 写死头注释 / Origin is legal, theta=0
        ELSE
            fXn := fX / fMaxC;                        // 归一 X / Normalised X
            fYn := fY / fMaxC;                        // 归一 Y / Normalised Y
            fA  := fMaxC * SQRT(fXn * fXn + fYn * fYn); // 归一后半径还原 / Radius restored after normalising
            fRad := ATAN2(fY, fX);                    // 反正切主值 [rad] / Principal arctangent [rad]
            fDeg := fRad * DL_POL_DEG180 / DL_POL_PI; // 换算角度 [deg] / Convert to degrees
            IF fDeg < 0.0 THEN
                fDeg := fDeg + 360.0;                 // 负角归入 0..360 / Wrap negative into 0..360
            END_IF
            IF fDeg >= 360.0 THEN
                fDeg := fDeg - 360.0;                 // 360 边界归一 / Normalise 360 boundary
            END_IF
            fB := fDeg;                               // 角度输出 [deg] / Angle output [deg]
        END_IF
        bValid := TRUE;                               // 正变换成立 / Forward transform valid
    eToCart:
        IF fX < 0.0 THEN
            uErrorId := 16#0001_0093;                 // 信息级：负半径语义歧义拒绝 / Info: negative radius rejected
            RETURN;                                   // 拒绝出口 / Rejection exit
        END_IF
        IF ABS(fY) > DL_POL_ANGMAX THEN
            fDeg := fY - 360.0 * TRUNC(fY / 360.0);   // 超域大角先取模防精度损失 / Huge angle reduced by modulo
            uErrorId := 16#0001_0094;                 // 信息级：角度超域已归一 / Info: angle out of range, normalised
        ELSE
            fDeg := fY;                               // 常规角原值生效 / Normal angle as-is
        END_IF
        fDeg := fDeg - 360.0 * TRUNC(fDeg / 360.0);   // 统一取模归一 / Uniform modulo normalisation
        IF fDeg < 0.0 THEN
            fDeg := fDeg + 360.0;                     // 取模后负值回正 / Wrap residual negative
        END_IF
        fRad := fDeg * DL_POL_PI / DL_POL_DEG180;     // 角度换算 [rad] / Convert to radians
        fA := fX * COS(fRad);                         // X = r·cos(theta) / X from radius and angle
        fB := fX * SIN(fRad);                         // Y = r·sin(theta) / Y from radius and angle
        bValid := TRUE;                               // 逆变换成立 / Inverse transform valid
    ELSE
        uErrorId := 16#0001_0095;                     // 信息级：模式非法兜底拒绝 / Info: illegal mode fallback
        RETURN;                                       // 拒绝出口 / Rejection exit
END_CASE
END_FUNCTION

(* ---- FC_DL_PowerUnitConvert.st ---- *)
(*==============================================================================
 * 组件名称 (Component)  : FC_DL_PowerUnitConvert
 * 所属子库 (Sublibrary) : DL_MathData
 * 当前版本 (Version)    : 1.0.0
 * 兼容性   (Platform)   : CODESYS 3.5+ / TwinCAT 3 / 汇川 InoProShop / 施耐德 Machine Expert
 *                         仅依赖 IEC 61131-3 算术运算符，零厂商私有库
 * 功能描述 (Function)   : 功率单位换算（系数表驱动）：以千瓦（kW）为中介单位，
 *                         fHub = fValue × kSrc，fResult = fHub ÷ kDst；系数为编译期
 *                         非零常量，纯常量除法，结构性无除零。
 *                         **符号语义**：功率允许负值（电动/发电四象限、能量回馈），
 *                         故本件**不做负值拒绝**，仅在结果非有限时兜底。
 *                         口径：HP 取机械马力（mechanical horsepower = 745.6998715822702 W），
 *                         非公制马力（735.49875 W）；两者差 1.4%，已在枚举注释中显式标定。
 * 接口     (Interface)  : 输入 fValue 被换算功率 [源单位]、eSrc 源单位、eDst 目标单位；
 *                         输出 fConverted 换算结果 [目标单位]、eErrCode（E_DL_PowerConvErr）；
 *                         返回值 = bValid 数值可信标志（TRUE = fConverted 可信）。
 * 边界     (Boundary)   : ① 属主边界：只做单位换算，不做功率因数修正、不做有功/无功分解。
 *                         ② 单位枚举越域 → 故障级 eInvalidUnit，结果哨兵 0。
 *                         ③ 非有限双判，命中即故障级 eNonFinite。
 *                         ④ 负值合法（回馈 / 发电象限），不置任何码。
 *                         ⑤ 零值 → 信息级 eZeroValue。
 *                         ⑥ kW ↔ W 跨越 1000 倍，结果复检防非有限。
 *                         ⑦ 零全局耦合（无 GVL / VAR_EXTERNAL / 物理地址）。
 * 分工声明 (Scope)      : 与 `FC_DL_EnergyUnitConvert` 分工：能量归那件；功率 × 时间 = 能量
 *                         的积分由调用方按时基完成（本件不持有时间量）。
 * 来源标签 (Source Tag) : 开源溯源：lgf-math 换算系数（公开物理常数，clean-room 重写）；许可证 MIT（仅参考语义，代码原创）
 * 码表     (Codes)      : 本件不占用全局数字码位；出口为 BOOL + LREAL +
 *                         本文件内定义 enum E_DL_PowerConvErr（全库唯一）。
 * 红线自检 (Redline)    : R1 ✓ 零 GVL/VAR_EXTERNAL ｜ R2 ✓ 零 %I/%Q/%M ｜ R3 ✓ 纯 IEC 61131-3
 *                         R4 ✓ 非有限双判 + 枚举域闸 + 常量除法无除零（负值按量纲放行） ｜ R5 ✓ 声明逐行同行双语注释
 *                         R6 N/A（纯函数无状态机） ｜ R7 N/A（无实例调用）
 * 修订历史 (Revision)   : 2026-11-23  v1.0.0  R77 首版（批次 B2 · 序号 18）
 * 验收向量 (Acceptance) : ① fValue=1.0, eSrc=eHp, eDst=eKw → 1×0.7456998715822702 = 0.7456998715822702 kW；
 *                         ② fValue=1.0, eSrc=eKw, eDst=eW → 1×1.0 = 1 kW, ÷0.001 = 1000.0 W；
 *                         ③ fValue=745.6998715822702, eSrc=eW, eDst=eHp → 0.7456998715822702 kW,
 *                         ÷0.7456998715822702 = 1.0 HP（容差 1E-12）；
 *                         ④ fValue=-11.0, eSrc=eKw, eDst=eW → -11000.0 W（负值合法）, eOk, TRUE；
 *                         ⑤ fValue=0.0, eSrc=eKw, eDst=eHp → 0.0, 返回 TRUE, eZeroValue。
 *==============================================================================*)

(*-----------------------------------------------------------------------------
 * 枚举: E_DL_PowerUnit（功率单位表，归属 DL_MathData，与本件同文件，全库唯一属主）
 *----------------------------------------------------------------------------*)
TYPE E_DL_PowerUnit :
(
    eKw := 0,   // 千瓦（中介单位） / Kilowatt, hub unit
    eHp := 1,   // 机械马力（= 0.7456998715822702 kW） / Mechanical horsepower
    eW  := 2    // 瓦（= 0.001 kW） / Watt
);
END_TYPE

(*-----------------------------------------------------------------------------
 * 枚举: E_DL_PowerConvErr（功率换算错误码）
 * 分级: 本件无「负值」故障码——功率负值属合法物理语义（回馈/发电）。
 *----------------------------------------------------------------------------*)
TYPE E_DL_PowerConvErr :
(
    eOk          := 0,   // 信息级：换算完成 / Info: conversion completed
    eZeroValue   := 1,   // 信息级：输入为零（合法） / Info: zero input, legal
    eInvalidUnit := 2,   // 故障级：单位枚举越域 / Fault: unit enum out of domain
    eNonFinite   := 3    // 故障级：输入非有限 / Fault: non-finite input
);
END_TYPE

FUNCTION FC_DL_PowerUnitConvert : BOOL
VAR_INPUT
    fValue : LREAL;           // 被换算功率值（可负） [源单位] / Power value, negative allowed, in source unit
    eSrc   : E_DL_PowerUnit;  // 源单位枚举 [-] / Source unit enum
    eDst   : E_DL_PowerUnit;  // 目标单位枚举 [-] / Destination unit enum
END_VAR
VAR_OUTPUT
    fConverted : LREAL;             // 换算结果（可负） [目标单位] / Converted result, may be negative
    eErrCode   : E_DL_PowerConvErr; // 错误码出口 [-] / Error code outlet
END_VAR
VAR
    _bNonFin : BOOL;   // 输入非有限当拍标志 [-] / Non-finite input flag
    _fHub    : LREAL;  // 中介功率值 [kW] / Hub power value in kilowatts
END_VAR
VAR CONSTANT
    DL_PUC2_KW   : LREAL := 1.0;                  // kW → kW 恒等系数 [-] / Hub identity factor
    DL_PUC2_HP   : LREAL := 0.7456998715822702;   // HP → kW 换算系数 [kW/HP] / Mechanical horsepower factor
    DL_PUC2_W    : LREAL := 0.001;                // W → kW 换算系数 [kW/W] / Watt factor
    DL_PUC2_ZERO : LREAL := 0.0;                  // 零值与非有限判零基准 [-] / Zero and non-finite base
END_VAR

(* —— 段 0：出口预置安全值 —— *)
FC_DL_PowerUnitConvert := FALSE;                   // 返回值预置无效 / Return preset invalid
fConverted := DL_PUC2_ZERO;                        // 结果哨兵 0 / Result sentinel
eErrCode   := E_DL_PowerConvErr.eInvalidUnit;      // 预置最严码 / Preset strictest code

(* —— 段 1：非有限域闸（R79 双判） —— *)
_bNonFin := (fValue <> fValue) OR ((fValue - fValue) <> DL_PUC2_ZERO);   // 非有限判定 / Non-finite test
IF _bNonFin THEN
    eErrCode := E_DL_PowerConvErr.eNonFinite;      // 故障级码 / Fault-level code
    RETURN;
END_IF

(* —— 段 2：极性说明（功率负值合法，本段仅注释占位，不做拦截） —— *)
(* Negative power is physically legal (regenerative quadrant), so no polarity gate is applied. *)

(* —— 段 3：源单位 → 中介 kW —— *)
IF eSrc = E_DL_PowerUnit.eKw THEN
    _fHub := fValue * DL_PUC2_KW;                  // 直通 / Hub pass-through
ELSIF eSrc = E_DL_PowerUnit.eHp THEN
    _fHub := fValue * DL_PUC2_HP;                  // HP × 0.7456998715822702 / Horsepower scaled
ELSIF eSrc = E_DL_PowerUnit.eW THEN
    _fHub := fValue * DL_PUC2_W;                   // W × 0.001 / Watt scaled
ELSE
    RETURN;                                        // 源单位越域 / Source unit out of domain
END_IF

(* —— 段 4：中介 kW → 目标单位（常量除法，分母非零） —— *)
IF eDst = E_DL_PowerUnit.eKw THEN
    fConverted := _fHub / DL_PUC2_KW;              // ÷1 / Divide by identity
ELSIF eDst = E_DL_PowerUnit.eHp THEN
    fConverted := _fHub / DL_PUC2_HP;              // ÷0.7456998715822702 / Divide by horsepower factor
ELSIF eDst = E_DL_PowerUnit.eW THEN
    fConverted := _fHub / DL_PUC2_W;               // ÷0.001 / Divide by watt factor
ELSE
    eErrCode   := E_DL_PowerConvErr.eInvalidUnit;  // 目标单位越域 / Destination out of domain
    fConverted := DL_PUC2_ZERO;
    RETURN;
END_IF

(* —— 段 5：结果非有限复检兜底 —— *)
IF (fConverted <> fConverted) OR ((fConverted - fConverted) <> DL_PUC2_ZERO) THEN
    fConverted := DL_PUC2_ZERO;                    // 复检异常回哨兵 / Recheck failed: sentinel
    eErrCode   := E_DL_PowerConvErr.eNonFinite;    // 故障级码 / Fault-level code
    RETURN;
END_IF

(* —— 段 6：成功出口 —— *)
IF fValue = DL_PUC2_ZERO THEN
    eErrCode := E_DL_PowerConvErr.eZeroValue;      // 信息级：零值 / Info: zero value
ELSE
    eErrCode := E_DL_PowerConvErr.eOk;             // 信息级成功 / Info success
END_IF
FC_DL_PowerUnitConvert := TRUE;                    // 换算有效 / Conversion valid

END_FUNCTION

(* ---- FC_DL_PressUnitConvert.st ---- *)
(*==============================================================================
 * 组件名称 (Component)  : FC_DL_PressUnitConvert
 * 所属子库 (Sublibrary) : DL_MathData
 * 当前版本 (Version)    : 1.0.0
 * 兼容性   (Platform)   : CODESYS 3.5+ / TwinCAT 3 / 汇川 InoProShop / 施耐德 Machine Expert
 *                         仅依赖 Standard.library（ABS），零厂商私有库
 * 功能描述 (Function)   : 压力工程量单位换算（系数表驱动）：以 Pa 为中介单位，
 *                         fPaAbs = fValue × kSrc，fResult = fPaAbs ÷ kDst，
 *                         kSrc/kDst 取自本文件常量系数表（纯常量除法，分母为非零
 *                         字面常量，结构性无除零）。负压域合法（表压/真空侧负读数
 *                         允许换算），换算结果落在绝对真空下限（0 Pa）之下时钳位
 *                         至 0 并置信息码 eClampVacuum（量值方向可饱和，规格指定）。
 *                         非有限输入 → 故障码 eNonFinite，输出哨兵 0。
 * 接口     (Interface)  : 输入 fValue 被换算压力值（Pa 域口径，含负压）[Pa]、
 *                         eSrc 源单位枚举、eDst 目标单位枚举；
 *                         输出 fConverted 换算结果（钳位后）[目标单位]、
 *                         eErrCode 错误码（E_DL_PressConvErr）、
 *                         返回值 = 换算有效标志（BOOL，TRUE = 数值可信）。
 * 边界     (Boundary)   : ① **属主边界（写死）：本件只做单位换算，不做量程标定、
 *                         不做表压/绝压模式判别**（调用方自行决定口径后传入）。
 *                         ② eSrc/eDst 超出枚举合法域（<0 或 >eMmHg）→ 故障码
 *                         eInvalidUnit，输出哨兵 0（ENUM 强转越域防御）。
 *                         ③ 系数表五个系数均为非零编译期常量，除法分母结构性
 *                         非零，无除零路径。
 *                         ④ 非有限判据：NaN 用自反 x <> x，Inf 用 (x−x) <> (x−x)
 *                         （R79 双判，无裸近似阈值）。
 *                         ⑤ 真空下限钳位只钳下限不设上限（量值饱和单向，正解
 *                         方向故障级码不启用，信息级 eClampVacuum 不置 bError）。
 *                         ⑥ 零全局耦合（无 GVL / VAR_EXTERNAL / 物理地址）。
 * 分工声明 (Scope)      : 与 `FB_DL_AnalogTransmitter` 分工：原始量程标定归那件、
 *                         工程量单位间换算归本件；本件不调用任何 FB，纯函数。
 * 来源标签 (Source Tag) : 自研线（SI 换算系数为公开物理常数定义，clean-room）
 * 码表     (Codes)      : 本件不占用任何全局数字码位。出口为 BOOL 返回 +
 *                         LREAL 结果 + ENUM eErrCode（本文件内定义，全库唯一）；
 *                         数字码位待主控收口阶段统一派号。
 * 红线自检 (Redline)    : R1 ✓ 零 GVL/VAR_EXTERNAL ｜ R2 ✓ 零 %I/%Q/%M ｜ R3 ✓ 纯 IEC 61131-3
 *                         R4 ✓ 非有限双判 + 单位域闸 + 真空下限钳位 ｜ R5 ✓ 声明逐行同行双语注释
 *                         R6 N/A（纯函数无状态机） ｜ R7 N/A（无实例调用）
 * 修订历史 (Revision)   : 2026-11-20  v1.0.0  R50 首版（批次 1 · 序号 1）
 * 验收向量 (Acceptance) : ① fValue=1.0, eSrc=eBar, eDst=ePa → 1×100000÷1
 *                         = 100000.0 Pa，返回 TRUE，eErrCode=eOk；
 *                         ② fValue=14.6959488, eSrc=ePsi, eDst=eBar →
 *                         14.6959488×6894.757293168761 ≈ 101325.0 Pa，
 *                         ÷100000 ≈ 1.01325 bar（容差 1E-6），eOk；
 *                         ③ fValue=760.0, eSrc=eMmHg, eDst=eKpa →
 *                         760×133.322387415 ≈ 101325.014 Pa，÷1000
 *                         ≈ 101.325014 kPa，eOk；
 *                         ④ fValue=-50000.0, eSrc=ePa, eDst=ePa → 中介值
 *                         <0 钳 0，输出 0.0，返回 TRUE，eErrCode=eClampVacuum
 *                         （信息级，bError 不置）。
 *==============================================================================*)

(*-----------------------------------------------------------------------------
 * 枚举: E_DL_PressUnit（压力单位表，归属 DL_MathData，与 FC_DL_PressUnitConvert
 *       同文件，全库唯一属主）
 *----------------------------------------------------------------------------*)
TYPE E_DL_PressUnit :
(
    ePa    := 0,   // 帕斯卡（中介单位） / Pascal, hub unit
    eKpa   := 1,   // 千帕 / Kilopascal
    eBar   := 2,   // 巴 / Bar
    ePsi   := 3,   // 磅每平方英寸 / Pound per square inch
    eMmHg  := 4    // 毫米汞柱（0 ℃ 托） / Millimetre of mercury at 0 degC
);
END_TYPE

(*-----------------------------------------------------------------------------
 * 枚举: E_DL_PressConvErr（错误码，故障级置 bError，信息级不置）
 *----------------------------------------------------------------------------*)
TYPE E_DL_PressConvErr :
(
    eOk          := 0,   // 成功 / Success
    eInvalidUnit := 1,   // 故障级：源/目标单位枚举越域 / Fault: unit enum out of domain
    eNonFinite   := 2,   // 故障级：输入非有限（NaN/Inf） / Fault: non-finite input
    eClampVacuum := 3    // 信息级：低于绝对真空下限已钳 0 / Info: clamped to absolute vacuum floor
);
END_TYPE

FUNCTION FC_DL_PressUnitConvert : BOOL
VAR_INPUT
    fValue   : LREAL;                 // 被换算压力值（负压域合法） [Pa] / Input pressure value, negative domain legal [Pa]
    eSrc     : E_DL_PressUnit;        // 源单位枚举 [-] / Source unit enum
    eDst     : E_DL_PressUnit;        // 目标单位枚举 [-] / Destination unit enum
END_VAR
VAR_OUTPUT
    fConverted : LREAL;               // 换算结果（真空下限钳位后） [目标单位] / Converted result after vacuum floor clamp
    eErrCode   : E_DL_PressConvErr;   // 错误码出口 / Error code outlet
END_VAR
VAR
    _bNonFin  : BOOL;                 // 输入非有限当拍量 [-] / Non-finite input flag
    _fPaAbs   : LREAL;                // 中介绝对压力值 [Pa] / Hub absolute pressure value
END_VAR
VAR CONSTANT
    DL_PUC_KPA    : LREAL := 1000.0;              // kPa → Pa 换算系数 [Pa/kPa] / kPa to Pa factor
    DL_PUC_BAR    : LREAL := 100000.0;            // bar → Pa 换算系数 [Pa/bar] / bar to Pa factor
    DL_PUC_PSI    : LREAL := 6894.757293168761;   // psi → Pa 换算系数（15 位有效数字） [Pa/psi] / psi to Pa factor
    DL_PUC_MMHG   : LREAL := 133.322387415;       // mmHg(0℃) → Pa 换算系数 [Pa/mmHg] / mmHg to Pa factor
    DL_PUC_ONE    : LREAL := 1.0;                 // Pa → Pa 恒等系数 [Pa/Pa] / Pa identity factor
    DL_PUC_ZERO   : LREAL := 0.0;                 // 真空下限与非有限判零基准 [Pa] / Vacuum floor and non-finite zero base
    DL_PUC_UNITMAX: INT   := 4;                   // 枚举合法域上限（eMmHg） [-] / Unit enum domain ceiling
END_VAR

(* —— 段 0：出口预置安全值（四段式第一段：预置） —— *)
FC_DL_PressUnitConvert := FALSE;                  // 返回值预置无效 / Return preset invalid
fConverted := DL_PUC_ZERO;                        // 结果哨兵 0 / Result sentinel zero
eErrCode := E_DL_PressConvErr.eInvalidUnit;       // 预置最严码，域闸命中直接早退 / Preset strictest code

(* —— 段 1：非有限域闸（R79 双判：NaN 自反 + Inf 差自减） —— *)
_bNonFin := (fValue <> fValue) OR ((fValue - fValue) <> DL_PUC_ZERO);   // 非有限判定 / Non-finite test
IF _bNonFin THEN
    eErrCode := E_DL_PressConvErr.eNonFinite;     // 故障级码（R45 配对见段 6） / Fault code
    RETURN;                                       // 早退保持哨兵输出 / Early exit with sentinel
END_IF

(* —— 段 2：单位枚举域闸（按枚举成员逐值比较，不依赖平台 ENUM→INT 强转方言） —— *)
(* 按枚举成员逐值比较，避免依赖平台 ENUM→INT 强转方言 *)
IF (eSrc = E_DL_PressUnit.ePa) THEN
    _fPaAbs := fValue * DL_PUC_ONE;               // Pa 直通 / Pa pass-through
ELSIF (eSrc = E_DL_PressUnit.eKpa) THEN
    _fPaAbs := fValue * DL_PUC_KPA;               // kPa × 1000 / kPa scaled
ELSIF (eSrc = E_DL_PressUnit.eBar) THEN
    _fPaAbs := fValue * DL_PUC_BAR;               // bar × 100000 / bar scaled
ELSIF (eSrc = E_DL_PressUnit.ePsi) THEN
    _fPaAbs := fValue * DL_PUC_PSI;               // psi × 6894.757... / psi scaled
ELSIF (eSrc = E_DL_PressUnit.eMmHg) THEN
    _fPaAbs := fValue * DL_PUC_MMHG;              // mmHg × 133.322... / mmHg scaled
ELSE
    RETURN;                                       // 源单位越域：保持预置故障码与哨兵 0 / Source unit out of domain
END_IF

(* —— 段 3：真空下限钳位（负压域合法，仅钳绝对真空以下） —— *)
eErrCode := E_DL_PressConvErr.eOk;                // 预置成功 / Preset success
IF _fPaAbs < DL_PUC_ZERO THEN
    _fPaAbs := DL_PUC_ZERO;                       // 钳至绝对真空下限 / Clamp to vacuum floor
    eErrCode := E_DL_PressConvErr.eClampVacuum;   // 信息级（不置 bError，规格⑤） / Info-level code
END_IF

(* —— 段 4：目标单位反换算（常量除法，分母非零结构性无除零） —— *)
IF (eDst = E_DL_PressUnit.ePa) THEN
    fConverted := _fPaAbs / DL_PUC_ONE;           // ÷1 直通 / Divide by one
ELSIF (eDst = E_DL_PressUnit.eKpa) THEN
    fConverted := _fPaAbs / DL_PUC_KPA;           // ÷1000 / Divide by kPa factor
ELSIF (eDst = E_DL_PressUnit.eBar) THEN
    fConverted := _fPaAbs / DL_PUC_BAR;           // ÷100000 / Divide by bar factor
ELSIF (eDst = E_DL_PressUnit.ePsi) THEN
    fConverted := _fPaAbs / DL_PUC_PSI;           // ÷6894.757... / Divide by psi factor
ELSIF (eDst = E_DL_PressUnit.eMmHg) THEN
    fConverted := _fPaAbs / DL_PUC_MMHG;          // ÷133.322... / Divide by mmHg factor
ELSE
    eErrCode := E_DL_PressConvErr.eInvalidUnit;   // 目标单位越域：回置故障码 / Destination unit out of domain
    fConverted := DL_PUC_ZERO;                    // 结果回哨兵 0 / Result back to sentinel
    RETURN;                                       // 早退 / Early exit
END_IF

(* —— 段 5：结果非有限复检兜底（四段式第四段：复检） —— *)
IF (_fPaAbs <> _fPaAbs) OR ((_fPaAbs - _fPaAbs) <> DL_PUC_ZERO) THEN
    fConverted := DL_PUC_ZERO;                    // 中介值复检异常：回哨兵 / Hub recheck failed: sentinel
    eErrCode := E_DL_PressConvErr.eNonFinite;     // 故障级码 / Fault code
    RETURN;                                       // 早退 / Early exit
END_IF

(* —— 段 6：成功出口（bError 由调用方按 eErrCode 归约；故障级码恒伴返回 FALSE） —— *)
FC_DL_PressUnitConvert := TRUE;                   // 换算有效（信息级钳位也算有效换算） / Conversion valid

END_FUNCTION

(* ---- FC_DL_PressureAltitudeCalc.st ---- *)
//==============================================================================
// 函数：FC_DL_PressureAltitudeCalc ｜ 中文名称：ISA 标准大气气压↔海拔双向换算
// 所属子库：DL_MathData ｜ 版本：v1.0.1 ｜ 日期：2026-11-23
// 兼容：CODESYS V3.5+ / TwinCAT 3 / 汇川 InoProShop / Machine Expert（纯标准库）
// 功能描述：ISA 对流层（0~11 km）标准大气双向换算。正解（海拔→气压）：
//           p = p0·(1 − L·h/T0)^(g/(R·L))；反解（气压→海拔）：
//           h = (T0/L)·(1 − (p/p0)^(R·L/g))。常量取 ISA 公开口径：
//           p0 = 101325 Pa、T0 = 288.15 K、L = 0.0065 K/m、
//           g = 9.80665 m/s2、R = 287.05287 J/(kg·K)。
// 开源溯源 (Origin)：原创实现（t1-2-oscat-building 建筑环境语义借用，ISA
//           公开公式，零外部源码行，clean-room 独立编写）
// 公开接口清单：输入 eMode / fValue；输出 fResult / bValid
// 错误码表：纯函数无状态机码轨；无效输入经 bValid = FALSE 表达（哨兵返回
//           0.0），本件不占用 16#0001 段码位（邻件免让位）
// 状态机：E_DL_PressAltMode（本文件唯一定义，全库唯一属主）：
//           eAltToPress = 0 / ePressToAlt = 1；枚举非法值走 CASE ELSE 兜底
// 边界行为：① 海拔域 [-500, 11000] m（ISA 对流层有效域，域外不外推）；
//           ② 气压域 [22632, 107477.5] Pa（对流层两端标准值，域外不外推；
//             −500 m 端值 R73 按公式订正）；
//           ③ L 恒非零为 ISA 常量，仍按纪律做非零断言常量（编译期保护）；
//           ④ 非有限输入（NaN 自反判 + 幅值判）→ 哨兵 0.0 返回；
//           ⑤ 枚举非法值 → CASE ELSE 哨兵返回。
// 修订历史：v1.0.0 2026-11-23 首版（R73 派单 · 批 2 · 序 8）
//           v1.0.1 2026-11-23 R73 返修：DL_PA_PMAX 按 ISA 标准大气公式订正
//           为 −500 m 对应值 107477.5 Pa（原 108900.0 与公式不符），边界
//           行为②同步订正。
//==============================================================================

(*------------------------------------------------------------------------------
 * 枚举: E_DL_PressAltMode（归属本函数，同文件发布，全库唯一属主）
 * 含义: 换算方向选择，成员与 CASE 标签双向完备。
 *-----------------------------------------------------------------------------*)
TYPE E_DL_PressAltMode :
(
    eAltToPress  := 0,  // 正解：输入海拔 [米]，输出气压 [帕] / Forward: altitude in, pressure out
    ePressToAlt  := 1   // 反解：输入气压 [帕]，输出海拔 [米] / Inverse: pressure in, altitude out
);
END_TYPE

(*------------------------------------------------------------------------------
 * 调用示例：fP := FC_DL_PressureAltitudeCalc(
 *             eMode := E_DL_PressAltMode.eAltToPress, fValue := 1500.0,
 *             bValid => bOk);
 * 注意：仅当 bValid = TRUE 时结果可进入判据；域外输入拒绝不外推。
 *-----------------------------------------------------------------------------*)
FUNCTION FC_DL_PressureAltitudeCalc : LREAL
VAR_INPUT
    eMode    : E_DL_PressAltMode;      // 换算方向枚举 [—] / Conversion direction enum
    fValue   : LREAL;                  // 输入量：海拔 [米] 或气压 [帕]，按 eMode 解释 / Input value, altitude [m] or pressure [Pa] per eMode
END_VAR
VAR_OUTPUT
    bValid   : BOOL;                   // 结果有效标志，FALSE 时返回哨兵 0.0 / Result validity flag
END_VAR
VAR CONSTANT
    DL_PA_P0   : LREAL := 101325.0;    // 海平面标准气压 [帕] / ISA sea-level standard pressure [Pa]
    DL_PA_T0   : LREAL := 288.15;      // 海平面标准温度 [开尔文] / ISA sea-level standard temperature [K]
    DL_PA_L    : LREAL := 0.0065;      // 对流层温度直减率 [开尔文每米] / ISA tropospheric lapse rate [K per m]
    DL_PA_G    : LREAL := 9.80665;     // 标准重力加速度 [米每平方秒] / Standard gravity [m per s2]
    DL_PA_R    : LREAL := 287.05287;   // 干空气气体常数 [焦每千克每开尔文] / Dry-air gas constant [J per kg per K]
    DL_PA_HMIN : LREAL := -500.0;      // 海拔有效下限 [米]（域外不外推）/ Altitude valid floor [m], no extrapolation
    DL_PA_HMAX : LREAL := 11000.0;     // 海拔有效上限 [米]（对流层顶）/ Altitude valid ceiling [m], tropopause
    DL_PA_PMIN : LREAL := 22632.0;     // 气压有效下限 [帕]（11 km 标准值）/ Pressure valid floor [Pa], 11 km ISA value
    DL_PA_PMAX : LREAL := 107477.5;    // 气压有效上限 [帕]（-500 m ISA 标准值，R73 订正：原 108900.0 与公式不符）/ Pressure valid ceiling [Pa], ISA value at -500 m, corrected
    DL_PA_EXP1 : LREAL := 5.2558797;   // 正解指数 g/(R·L) 预算值 [1] / Forward exponent g/(R*L), precomputed
    DL_PA_EXP2 : LREAL := 0.190263236; // 反解指数 R·L/g 预算值 [1] / Inverse exponent R*L/g, precomputed
    DL_PA_INF  : LREAL := 1.7976931348623157E308; // LREAL 幅值上限 / LREAL magnitude ceiling
    DL_PA_ZERO : LREAL := 0.0;         // 无效哨兵返回值 / Sentinel return for invalid
END_VAR

// ---- 段 1｜出口默认值（纯函数无实例，无定时器/沿刷新义务）----
bValid := FALSE;                      // 缺省无效 / Invalid by default

// ---- 段 2｜输入防御：非有限值（NaN 自反判 + Inf 幅值判，R79）----
IF (fValue <> fValue) OR (ABS(fValue) > DL_PA_INF) THEN
    FC_DL_PressureAltitudeCalc := DL_PA_ZERO; // 无效输入：哨兵零返回 / Invalid input, sentinel zero return
    RETURN;                            // 结构早退 / early exit
END_IF

// ---- 段 3｜双向换算主体（CASE 带 ELSE；域闸拒绝不外推）----
CASE eMode OF
    E_DL_PressAltMode.eAltToPress:     // 正解：海拔 → 气压
        IF (fValue < DL_PA_HMIN) OR (fValue > DL_PA_HMAX) THEN
            FC_DL_PressureAltitudeCalc := DL_PA_ZERO; // 海拔域外拒绝（哨兵零）/ Altitude out of range, refused
            RETURN;                    // 结构早退 / early exit
        END_IF
        FC_DL_PressureAltitudeCalc := DL_PA_P0
            * EXPT((1.0 - DL_PA_L * fValue / DL_PA_T0), DL_PA_EXP1); // 标准大气压 [帕] / ISA standard pressure [Pa]

    E_DL_PressAltMode.ePressToAlt:     // 反解：气压 → 海拔
        IF (fValue < DL_PA_PMIN) OR (fValue > DL_PA_PMAX) THEN
            FC_DL_PressureAltitudeCalc := DL_PA_ZERO; // 气压域外拒绝（哨兵零）/ Pressure out of range, refused
            RETURN;                    // 结构早退 / early exit
        END_IF
        FC_DL_PressureAltitudeCalc := (DL_PA_T0 / DL_PA_L)
            * (1.0 - EXPT((fValue / DL_PA_P0), DL_PA_EXP2)); // 标准海拔 [米] / ISA standard altitude [m]

    ELSE                               // 枚举非法值兜底（R21：CASE 必带 ELSE）
        FC_DL_PressureAltitudeCalc := DL_PA_ZERO; // 非法枚举：哨兵零返回 / Illegal enum, sentinel zero return
        RETURN;                        // 结构早退 / early exit
END_CASE

bValid := TRUE;                       // 全部防御通过：结果有效 / Result valid
END_FUNCTION

(* ---- FC_DL_RampStepReal.st ---- *)
(*==============================================================================
 * 组件名称 (Component)  : FC_DL_RampStepReal
 * 所属子库 (Sublibrary) : DL_MathData ｜ 版本 (Version) : 1.0.0 ｜ 2026-11-23
 * 兼容性   (Platform)   : CODESYS 3.5+ / TwinCAT 3 / 汇川 InoProShop / 施耐德 Machine Expert
 *                         仅依赖 IEC 61131-3 算术运算符与 ABS，零厂商私有库
 * 功能描述 (Function)   : 固定步长爬坡（FC 形态，纯组合逻辑）：把当前值 fX 沿目标 fXTarget
 *                         方向每拍最多推进 fStep，剩余量不足一步时直接到达目标（无过冲）。
 *                         fStep ≤ 0 → 不爬坡，直接输出 fXTarget（开关量式跳变，信息级 eDirectJump）。
 *                         本件不持有跨拍状态：当前值由调用方以 fX 传入，故可重入、可多处例化。
 * 接口     (Interface)  : 输入 fX 当前值 [工程单位]、fXTarget 目标值 [工程单位]、
 *                         fStep 每拍最大步长，有效域 > 0 [工程单位/拍]；
 *                         输出 fY 爬坡后输出 [工程单位]、bArrived 到达标志（本拍已在目标上）、
 *                         eErrCode（E_DL_RampStepErr）；返回值 = 数值可信标志。
 * 边界     (Boundary)   : ① fStep ≤ 0 → 直通目标（信息级 eDirectJump，返回值 TRUE）。
 *                         ② 任一浮点入参非有限 → 故障级 eNonFinite，fY = 0 哨兵，返回 FALSE。
 *                         ③ 到达判定用容差 DL_RSTP_EPS（1E-6），禁浮点判等（R4）。
 *                         ④ 输出复检非有限 → 回退 fX 并报故障（保持上一有效当前值）。
 *                         ⑤ 零全局耦合（无 GVL / VAR_EXTERNAL / 物理地址）。
 * 码表     (Codes)      : 本件不占用全局数字码位（R297 零码位范式）；出口为 BOOL + REAL +
 *                         本文件内 enum E_DL_RampStepErr（全库唯一属主）。
 * 分工声明 (Scope)      : 带到达判定与跨周期驻留的斜坡发生器归 FB_DL_RampGenerator 与
 *                         FB_DL_RampSoakProfile；本件只做单拍步进决策，不积分、不驻留。
 * 归属     (Ownership)  : E_DL_RampStepErr 归属本文件（全库唯一属主，R264）。
 * 红线自检 (Redline)    : R1 ✓ 零 GVL ｜ R2 ✓ 零 %I/%Q ｜ R3 ✓ 纯 IEC ｜ R4 ✓ 非有限双判 +
 *                         容差比较 + 无除法 ｜ R5 ✓ 逐行同行双语注释 ｜ R6 N/A（纯函数）
 *                         R7 N/A（无实例调用）
 * 修订历史 (Revision)   : 2026-11-23  v1.0.0  R78-B2 首版
 * 验收向量 (Acceptance) :
 *   A1 fX=0.0, fXTarget=10.0, fStep=3.0 → fY=3.0, bArrived=FALSE, eStepping；
 *   A2 fX=8.5, fXTarget=10.0, fStep=3.0 → 剩余 1.5 < 3.0 → fY=10.0, bArrived=TRUE, eArrived；
 *   A3 fX=10.0, fXTarget=0.0, fStep=4.0 → fY=6.0（下行），eStepping；
 *   A4 fX=0.0, fXTarget=10.0, fStep=0.0 → fY=10.0, eDirectJump, 返回 TRUE；
 *   A5 fXTarget=NaN → fY=0.0, eNonFinite, 返回 FALSE。
 *============================================================================*)

(*-----------------------------------------------------------------------------
 * 枚举: E_DL_RampStepErr（步长爬坡出口码；信息级 = 0..9，故障级 = 10 起）
 *----------------------------------------------------------------------------*)
TYPE E_DL_RampStepErr :
(
    eArrived    := 0,   // 信息级：本拍已到达目标 / Info: target reached this scan
    eStepping   := 1,   // 信息级：本拍推进一个步长 / Info: one step advanced this scan
    eDirectJump := 2,   // 信息级：步长越域，直接跳变到目标 / Info: step out of domain, jumped to target
    eNonFinite  := 10   // 故障级：入参或结果非有限 / Fault: non-finite input or result
);
END_TYPE

FUNCTION FC_DL_RampStepReal : BOOL
VAR_INPUT
    fX       : REAL;   // 当前值（调用方持有的实际值）[工程单位] / Current value held by the caller in engineering unit
    fXTarget : REAL;   // 目标值 [工程单位] / Target value in engineering unit
    fStep    : REAL;   // 每拍最大步长，有效域 > 0 [工程单位/拍] / Max step per scan, valid domain > 0
END_VAR
VAR_OUTPUT
    fY       : REAL;              // 爬坡后输出 [工程单位] / Ramped output in engineering unit
    bArrived : BOOL;              // 到达标志：本拍输出已在目标容差内 [-] / Arrived flag within tolerance this scan
    eErrCode : E_DL_RampStepErr;   // 出口码 [-] / Outlet code
END_VAR
VAR
    _bBadX      : BOOL;   // fX 非有限标志 [-] / Non-finite flag of fX
    _bBadTarget : BOOL;   // fXTarget 非有限标志 [-] / Non-finite flag of fXTarget
    _bBadStep   : BOOL;   // fStep 非有限标志 [-] / Non-finite flag of fStep
    _fRemain    : REAL;   // 剩余量 = 目标 − 当前 [工程单位] / Remaining distance in engineering unit
    _fAbsRemain : REAL;   // 剩余量绝对值 [工程单位] / Absolute remaining distance
END_VAR
VAR CONSTANT
    DL_RSTP_ZERO : REAL := 0.0;     // 零基准与符号分界 [-] / Zero base and sign boundary
    DL_RSTP_EPS  : REAL := 1.0E-6;  // 到达判定容差 [-] / Arrival tolerance
END_VAR

(* —— 段 0：出口预置安全侧 —— *)
FC_DL_RampStepReal := FALSE;                         // 返回值预置不可信 / Return preset not trustworthy
fY       := DL_RSTP_ZERO;                            // 输出哨兵 0 / Output sentinel
bArrived := FALSE;                                   // 到达标志预清（单拍位统一预置）/ Single-shot flag preset
eErrCode := E_DL_RampStepErr.eNonFinite;             // 预置最严码 / Preset strictest code

(* —— 段 1：入参非有限闸（R272 全量枚举 fX / fXTarget / fStep） —— *)
_bBadX      := (fX <> fX) OR ((fX - fX) <> DL_RSTP_ZERO);                    // 当前值非有限 / Current value non-finite
_bBadTarget := (fXTarget <> fXTarget) OR ((fXTarget - fXTarget) <> DL_RSTP_ZERO);  // 目标非有限 / Target non-finite
_bBadStep   := (fStep <> fStep) OR ((fStep - fStep) <> DL_RSTP_ZERO);        // 步长非有限 / Step non-finite
IF _bBadX OR _bBadTarget OR _bBadStep THEN
    RETURN;                                          // 故障出口：fY 保持 0 哨兵 / Fault exit, sentinel kept
END_IF

(* —— 段 2：步长域闸（fStep ≤ 0 → 不做爬坡，直接跳变到目标） —— *)
IF fStep <= DL_RSTP_ZERO THEN
    fY       := fXTarget;                            // 直通目标 / Jump straight to the target
    bArrived := TRUE;                                // 目标即到位 / Target equals arrival
    eErrCode := E_DL_RampStepErr.eDirectJump;        // 信息级：直接跳变 / Info: direct jump
    FC_DL_RampStepReal := TRUE;                      // 输出可信 / Output trustworthy
    RETURN;
END_IF

(* —— 段 3：剩余量与步进决策（不足一步即到达，结构性无过冲） —— *)
_fRemain    := fXTarget - fX;                        // 剩余量 / Remaining distance
_fAbsRemain := ABS(_fRemain);                        // 剩余量绝对值 / Absolute remaining distance
IF _fAbsRemain <= DL_RSTP_EPS THEN
    fY       := fXTarget;                            // 已在目标上：锁定目标 / Already there: lock the target
    bArrived := TRUE;                                // 到达标志 / Arrived flag
    eErrCode := E_DL_RampStepErr.eArrived;           // 信息级：已到达 / Info: arrived
ELSIF _fAbsRemain <= (fStep + DL_RSTP_EPS) THEN
    fY       := fXTarget;                            // 剩余不足一步：到达且不过冲 / Sub-step remainder: arrive without overshoot
    bArrived := TRUE;                                // 到达标志 / Arrived flag
    eErrCode := E_DL_RampStepErr.eArrived;           // 信息级：已到达 / Info: arrived
ELSE
    IF _fRemain > DL_RSTP_ZERO THEN
        fY := fX + fStep;                            // 上行推进一个步长 / Step upward
    ELSE
        fY := fX - fStep;                            // 下行推进一个步长 / Step downward
    END_IF
    bArrived := FALSE;                               // 未到达 / Not arrived
    eErrCode := E_DL_RampStepErr.eStepping;          // 信息级：推进中 / Info: stepping
END_IF

(* —— 段 4：结果复检（推进后非有限 → 回退当前值并报故障） —— *)
IF (fY <> fY) OR ((fY - fY) <> DL_RSTP_ZERO) THEN
    fY       := fX;                                  // 回退当前值 / Fall back to the current value
    bArrived := FALSE;                               // 到达标志撤销 / Arrival flag withdrawn
    eErrCode := E_DL_RampStepErr.eNonFinite;         // 故障级码 / Fault-level code
    FC_DL_RampStepReal := FALSE;                     // 故障出口不可信 / Fault exit not trustworthy
    RETURN;
END_IF

FC_DL_RampStepReal := TRUE;                          // 输出可信 / Output trustworthy
END_FUNCTION

(* ---- FC_DL_RateLimitReal.st ---- *)
(*==============================================================================
 * 组件名称 (Component)  : FC_DL_RateLimitReal
 * 所属子库 (Sublibrary) : DL_MathData ｜ 版本 (Version) : 1.0.0 ｜ 2026-11-23
 * 兼容性   (Platform)   : CODESYS 3.5+ / TwinCAT 3 / 汇川 InoProShop / 施耐德 Machine Expert
 *                         仅依赖 IEC 61131-3 算术运算符与 ABS，零厂商私有库
 * 功能描述 (Function)   : 单拍斜率限幅（FC 形态）：本拍原始输入 fX 与上一拍受限输出
 *                         fXPrev 之差超过 fRateMax × fDt 时，按最大步进逼近，否则直通。
 *                         **契约补充声明**：斜率限幅在数学上必须持有「上一拍输出」，
 *                         故本件使用 VAR_IN_OUT 引脚 fXPrev（调用方声明为静态变量），
 *                         首拍或 fXPrev 被污染时以本拍 fX 重建（置信息码 ePrevRebuilt）。
 *                         严格无内部状态，可重入、可多处例化。
 * 接口     (Interface)  : 输入 fX 原始输入 [工程单位]、fRateMax 限幅速率 [单位/秒]、
 *                         fDt 采样周期 [s]；VAR_IN_OUT fXPrev 上一拍受限输出（本件写回）；
 *                         输出 fY 限幅输出 [工程单位]、eErrCode（E_DL_RateLimitErr）；
 *                         返回值 = 数值可信标志（TRUE = fY 可信）。
 * 边界     (Boundary)   : ① fRateMax ≤ 0 或 fDt ≤ 0 → 旁路，fY = fX（信息级 eBypass，
 *                             返回值 TRUE——旁路输出仍是原值的忠实搬运，非故障）。
 *                         ② 任一浮点入参非有限（NaN / ±Inf）→ 故障级 eNonFinite，
 *                            fY = 0 哨兵，返回 FALSE（R79 双判，禁近似阈值）。
 *                         ③ 步进 fRateMax × fDt 溢出为非有限 → 同按旁路处理（不再逼近）。
 *                         ④ 限幅后结果复检，非有限则回退到 fXPrev 并报故障。
 *                         ⑤ 浮点同值比较一律用容差 DL_RLIM_EPS（1E-6），禁 `=`（R4）。
 *                         ⑥ 零全局耦合（无 GVL / VAR_EXTERNAL / 物理地址）。
 * 码表     (Codes)      : 本件不占用全局数字码位（R297 零码位范式）；出口为 BOOL +
 *                         REAL + 本文件内 enum E_DL_RateLimitErr（全库唯一属主）。
 *                         信息级码 eLimited / eBypass / ePrevRebuilt 永不置错；
 *                         故障级码 eNonFinite 伴随返回值 FALSE。
 * 分工声明 (Scope)      : 有状态斜坡发生（跨周期积分 + 到达标志）归 FB_DL_RampGenerator；
 *                         本件为纯函数形态单拍限幅，供扫描内计算链使用。
 * 归属     (Ownership)  : E_DL_RateLimitErr 归属本文件（全库唯一属主，R264）。
 * 红线自检 (Redline)    : R1 ✓ 零 GVL ｜ R2 ✓ 零 %I/%Q ｜ R3 ✓ 纯 IEC ｜ R4 ✓ 非有限双判 +
 *                         除零结构不可达（无除法）+ 容差比较 ｜ R5 ✓ 逐行同行双语注释
 *                         R6 N/A（纯函数无状态机） ｜ R7 N/A（无实例调用）
 * 修订历史 (Revision)   : 2026-11-23  v1.0.0  R78-B2 首版
 * 验收向量 (Acceptance) :
 *   A1 fX=10.0, fPrev=0.0, fRateMax=2.0, fDt=1.0 → 步进 2.0 → fY=2.0, eLimited；
 *   A2 续 A1：fX=10.0, fPrev=2.0, fRateMax=2.0, fDt=1.0 → fY=4.0, eLimited；
 *   A3 fX=3.0, fPrev=2.0, fRateMax=2.0, fDt=1.0 → 增量 1.0 ≤ 2.0 → fY=3.0, eOk；
 *   A4 fX=5.0, fPrev=2.0, fRateMax=0.0, fDt=1.0 → 旁路 → fY=5.0, eBypass, 返回 TRUE；
 *   A5 fX=NaN, fPrev=2.0 → fY=0.0, eNonFinite, 返回 FALSE。
 *============================================================================*)

(*-----------------------------------------------------------------------------
 * 枚举: E_DL_RateLimitErr（斜率限幅出口码；信息级 = 0..9，故障级 = 10 起）
 *----------------------------------------------------------------------------*)
TYPE E_DL_RateLimitErr :
(
    eOk          := 0,   // 信息级：未超速，直通 / Info: within rate, pass-through
    eLimited     := 1,   // 信息级：本拍已按最大步进逼近 / Info: closed in by the max step this scan
    eBypass      := 2,   // 信息级：速率或周期越域，旁路输出原值 / Info: rate or period out of domain, bypassed
    ePrevRebuilt := 3,   // 信息级：fXPrev 未初始化或被污染，已用本拍 fX 重建 / Info: previous output rebuilt from fX
    eNonFinite   := 10   // 故障级：入参或结果非有限 / Fault: non-finite input or result
);
END_TYPE

FUNCTION FC_DL_RateLimitReal : BOOL
VAR_INPUT
    fX       : REAL;   // 本拍原始输入 [工程单位] / Raw input this scan in engineering unit
    fRateMax : REAL;   // 允许最大变化速率，有效域 > 0 [单位/秒] / Max allowed rate, valid domain > 0 in unit per second
    fDt      : REAL;   // 采样周期，有效域 > 0 [s] / Sampling period, valid domain > 0 in seconds
END_VAR
VAR_IN_OUT
    fXPrev : REAL;     // 上一拍受限输出，本件写回新值 [工程单位] / Previous limited output, written back by this function
END_VAR
VAR_OUTPUT
    fY       : REAL;              // 限幅输出 [工程单位] / Rate-limited output in engineering unit
    eErrCode : E_DL_RateLimitErr;  // 出口码 [-] / Outlet code
END_VAR
VAR
    _bBadX     : BOOL;   // fX 非有限标志 [-] / Non-finite flag of fX
    _bBadRate  : BOOL;   // fRateMax 非有限标志 [-] / Non-finite flag of fRateMax
    _bBadDt    : BOOL;   // fDt 非有限标志 [-] / Non-finite flag of fDt
    _bBadPrev  : BOOL;   // fXPrev 非有限标志 [-] / Non-finite flag of fXPrev
    _fMaxStep  : REAL;   // 本拍允许最大步进 = fRateMax × fDt [工程单位] / Max step this scan
    _fDelta    : REAL;   // 原始增量 = fX − fXPrev [工程单位] / Raw delta between input and previous output
    _fAbsDelta : REAL;   // 增量绝对值 [工程单位] / Absolute delta
END_VAR
VAR CONSTANT
    DL_RLIM_ZERO : REAL := 0.0;     // 零基准与符号分界 [-] / Zero base and sign boundary
    DL_RLIM_EPS  : REAL := 1.0E-6;  // 浮点同值判定容差 [-] / Float equality tolerance
END_VAR

(* —— 段 0：出口预置安全侧 —— *)
FC_DL_RateLimitReal := FALSE;                        // 返回值预置不可信 / Return preset not trustworthy
fY      := DL_RLIM_ZERO;                             // 输出哨兵 0 / Output sentinel
eErrCode := E_DL_RateLimitErr.eNonFinite;            // 预置最严码 / Preset strictest code

(* —— 段 1：入参非有限闸（R272 全量枚举 fX / fRateMax / fDt） —— *)
_bBadX    := (fX <> fX) OR ((fX - fX) <> DL_RLIM_ZERO);                    // fX 非有限 / fX non-finite
_bBadRate := (fRateMax <> fRateMax) OR ((fRateMax - fRateMax) <> DL_RLIM_ZERO);  // 速率非有限 / Rate non-finite
_bBadDt   := (fDt <> fDt) OR ((fDt - fDt) <> DL_RLIM_ZERO);                // 周期非有限 / Period non-finite
IF _bBadX OR _bBadRate OR _bBadDt THEN
    RETURN;                                          // 故障出口：fY 保持 0 哨兵 / Fault exit, sentinel kept
END_IF

(* —— 段 2：上一拍输出有效性闸（未初始化或已被污染 → 用本拍输入重建，防 NaN 搬运） —— *)
_bBadPrev := (fXPrev <> fXPrev) OR ((fXPrev - fXPrev) <> DL_RLIM_ZERO);     // 前值非有限 / Previous value non-finite
IF _bBadPrev THEN
    fXPrev   := fX;                                  // 以本拍输入重建起点 / Rebuild the starting point
    eErrCode := E_DL_RateLimitErr.ePrevRebuilt;      // 信息级：前值已重建 / Info: previous value rebuilt
END_IF

(* —— 段 3：速率 / 周期域闸（fRateMax ≤ 0 或 fDt ≤ 0 → 旁路，输出原 x） —— *)
IF (fRateMax <= DL_RLIM_ZERO) OR (fDt <= DL_RLIM_ZERO) THEN
    fY      := fX;                                   // 旁路：输出保持原 x / Bypass: output keeps the raw input
    fXPrev  := fX;                                   // 前值同步 / Previous value follows
    eErrCode := E_DL_RateLimitErr.eBypass;           // 信息级：旁路 / Info: bypassed
    FC_DL_RateLimitReal := TRUE;                     // 旁路输出可信 / Bypass output is trustworthy
    RETURN;
END_IF

(* —— 段 4：本拍最大步进（乘后复检，溢出为非有限则旁路） —— *)
_fMaxStep := fRateMax * fDt;                         // 步进 = 速率 × 周期 / Step equals rate times period
IF (_fMaxStep <> _fMaxStep) OR ((_fMaxStep - _fMaxStep) <> DL_RLIM_ZERO) THEN
    fY      := fX;                                   // 步进不可表：放弃逼近 / Unrepresentable step: no approach
    fXPrev  := fX;                                   // 前值同步 / Previous value follows
    eErrCode := E_DL_RateLimitErr.eBypass;           // 信息级：旁路 / Info: bypassed
    FC_DL_RateLimitReal := TRUE;                     // 原值可信 / Raw value is trustworthy
    RETURN;
END_IF

(* —— 段 5：增量比较与逼近（超速按符号方向各逼近一步，方向分列 R146） —— *)
_fDelta    := fX - fXPrev;                           // 原始增量 / Raw delta
_fAbsDelta := ABS(_fDelta);                          // 增量绝对值 / Absolute delta
IF _fAbsDelta <= (_fMaxStep + DL_RLIM_EPS) THEN
    fY      := fX;                                   // 未超速：直通 / Within rate: pass-through
    eErrCode := E_DL_RateLimitErr.eOk;               // 信息级：正常 / Info: normal
ELSE
    IF _fDelta > DL_RLIM_ZERO THEN
        fY := fXPrev + _fMaxStep;                    // 上行逼近 / Approach upward
    ELSE
        fY := fXPrev - _fMaxStep;                    // 下行逼近 / Approach downward
    END_IF
    eErrCode := E_DL_RateLimitErr.eLimited;          // 信息级：本拍受限 / Info: limited this scan
END_IF

(* —— 段 6：结果复检（逼近后仍非有限 → 回退前值并报故障） —— *)
IF (fY <> fY) OR ((fY - fY) <> DL_RLIM_ZERO) THEN
    fY      := fXPrev;                               // 回退上一有效值 / Fall back to the last valid value
    eErrCode := E_DL_RateLimitErr.eNonFinite;        // 故障级码 / Fault-level code
    FC_DL_RateLimitReal := FALSE;                    // 故障出口不可信 / Fault exit not trustworthy
    RETURN;
END_IF

fXPrev := fY;                                        // 前值写回（唯一写入点）/ Single write-back point
FC_DL_RateLimitReal := TRUE;                         // 输出可信 / Output trustworthy
END_FUNCTION

(* ---- FC_DL_RtdLinearization.st ---- *)
(*
  ==================================================================
  组件名 Component  : FC_DL_RtdLinearization
  分类   Category   : DL_MathData
  复杂度 Complexity  : cx4
  版本   Version    : 1.0.0
  功能   Purpose    : Pt100 / Pt1000 阻值到温度的 Callendar-Van Dusen（CVD）反解。
                      T >= 0 段用二次方程求根公式；T < 0 段（含 C(T-100)T³ 项）
                      用定点迭代收敛反解。三线制引线电阻补偿先行扣除；R 越出
                      [R(-200C), R(850C)] 置 bOutOfRange（出口取安全侧零），非有限
                      或 R_eff <= 0 置 bInvalid。
  来源   Source     : ROADMAP R56 池 / T2 自研（IEC 60751 公开系数）
  溯源   Origin     : IEC 61131-3 标准语义的道莅防御性实现；CVD 方程与 A / B / C
                      系数为 IEC 60751 公开标准值，clean-room 自研实现，未复制任何
                      闭源代码行。
  平台   Platform   : 纯 IEC 61131-3（LREAL / SQRT，无私有库、无幂运算符）
  作者   Author     : 道莅代码库 · PLC 编程专家（R56）
  ------------------------------------------------------------------
  边界 Boundary     :
                      一 本件只做 RTD 阻值反解温度，不做单位换算、不做查表（属主边界）；
                      二 CVD 系数取 IEC 60751 标准值：R0(Pt100)=100 / R0(Pt1000)=1000，
                         A=3.9083E-3，B=-5.775E-7，C=-4.183E-12；
                      三 测温域 [-200, 850] 摄氏度，对应 Pt100 阻值域 [18.52, 390.48] 欧，
                         Pt1000 为其十倍；
                      四 负温段定点迭代收缩因子上界约 0.07（B·2T/A 在 T=-200 处），
                         60 次迭代含 1.0E-9 收敛阈足够；不收敛置 bInvalid；
                      五 无全局变量、无外部变量声明、无物理地址寻址、无定时器（纯函数）。
  输出契约 Output contract:
                      fTempC 仅在 bInvalid = FALSE 且 bOutOfRange = FALSE 时有效；
                      标志优先级 bInvalid > bOutOfRange；本件为纯函数，无跨扫描周期状态驻留。
  修订记录 Revision  :
    2026-11-20  v1.0.0  R56 首版（批 1 · 序号 4）
  ==================================================================
*)

TYPE E_DL_RtdType :
(
    ePt100  := 0, // Pt100 铂电阻，R0 = 100 欧 / Pt100 RTD with R0 of one hundred ohm
    ePt1000 := 1  // Pt1000 铂电阻，R0 = 1000 欧 / Pt1000 RTD with R0 of one thousand ohm
);
END_TYPE

FUNCTION FC_DL_RtdLinearization : BOOL
VAR_INPUT
    fROhm    : LREAL;        // RTD 实测阻值（含引线电阻）[欧] / measured RTD resistance including the leads [ohm]
    eType    : E_DL_RtdType; // RTD 类型选择 [枚举] / RTD type selector [enum]
    fLeadOhm : LREAL;        // 三线制引线电阻补偿量（从实测中扣除）[欧] / three wire lead resistance to be subtracted [ohm]
END_VAR
VAR_OUTPUT
    fTempC     : LREAL;      // 反解温度 [摄氏度] / solved temperature [degree celsius]
    bOutOfRange: BOOL;       // 阻值越出测温域 [-] / the resistance is outside the measuring domain
    bInvalid   : BOOL;       // 输入非有限或阻值无效 [-] / input non finite or the resistance void
END_VAR
VAR
    _bFin   : BOOL := FALSE;    // 两个实数输入全部有限 [-] / both real inputs are finite
    _fR0    : LREAL := 100.0;   // 标称零度阻值 [欧] / nominal resistance at zero degree [ohm]
    _fA     : LREAL := 3.9083E-3;   // CVD 一次系数 [每摄氏度] / CVD coefficient A [per degree celsius]
    _fB     : LREAL := -5.775E-7;   // CVD 二次系数 [每平方摄氏度] / CVD coefficient B [per square degree celsius]
    _fC     : LREAL := -4.183E-12;  // CVD 负温系数 [每四次摄氏度] / CVD coefficient C for the negative range [per fourth degree celsius]
    _fRMin  : LREAL := 18.52;   // 测温域下限阻值（-200 摄氏度）[欧] / domain floor resistance at minus two hundred [ohm]
    _fRMax  : LREAL := 390.48;  // 测温域上限阻值（850 摄氏度）[欧] / domain ceiling resistance at eight fifty [ohm]
    _fRUse  : LREAL := 0.0;     // 扣除引线后的有效阻值 [欧] / effective resistance after the lead subtraction [ohm]
    _fRel   : LREAL := 0.0;     // 相对阻值 R/R0 [无量纲] / relative resistance over R0
    _fDisc  : LREAL := 0.0;     // 二次方程判别式 [无量纲] / quadratic discriminant
    _fTPos  : LREAL := 0.0;     // 正温段求根结果 [摄氏度] / the positive branch root [degree celsius]
    _fTIt   : LREAL := 0.0;     // 负温段迭代值 [摄氏度] / the negative branch iterate [degree celsius]
    _fTNext : LREAL := 0.0;     // 负温段下个迭代值 [摄氏度] / the next negative branch iterate [degree celsius]
    _fDlt   : LREAL := 0.0;     // 迭代步差 [摄氏度] / the iterate step difference [degree celsius]
    _nI     : INT := 0;         // 迭代守护游标 [次] / iteration guard cursor [count]
    _bConv  : BOOL := FALSE;    // 迭代收敛标志 [-] / iteration convergence flag
END_VAR

// 段 1｜非有限闸（R151）与类型分派 / segment 1, finiteness gate and the type dispatch
_bFin := (fROhm = fROhm) AND ((fROhm - fROhm) = (fROhm - fROhm)) AND (fLeadOhm = fLeadOhm) AND ((fLeadOhm - fLeadOhm) = (fLeadOhm - fLeadOhm)); // 两实数输入有限性 / finiteness of both real inputs
bInvalid := NOT _bFin; // 非有限即无效 / non finite means invalid
bOutOfRange := FALSE; // 越域标志预置假 / preset the out of range flag to false
fTempC := 0.0; // 出口预置安全侧零（R127）/ preset the outlet to the safe side zero
CASE eType OF // 类型分派，常量在 CASE 内按型落定 / the type dispatch, the constants settle per type
E_DL_RtdType.ePt100: // Pt100 / the Pt100 type
    _fR0 := 100.0;   // 零度阻值 [欧] / the zero degree resistance [ohm]
    _fRMin := 18.52; // -200 摄氏度阻值下限 [欧] / the floor at minus two hundred [ohm]
    _fRMax := 390.48; // 850 摄氏度阻值上限 [欧] / the ceiling at eight fifty [ohm]
E_DL_RtdType.ePt1000: // Pt1000 / the Pt1000 type
    _fR0 := 1000.0;   // 零度阻值 [欧] / the zero degree resistance [ohm]
    _fRMin := 185.2;  // -200 摄氏度阻值下限 [欧] / the floor at minus two hundred [ohm]
    _fRMax := 3904.8; // 850 摄氏度阻值上限 [欧] / the ceiling at eight fifty [ohm]
ELSE // 非法类型枚举兜底（R128）/ the illegal type fallback
    bInvalid := TRUE; // 置无效标志 / raise the invalid flag
END_CASE
IF bInvalid THEN // 非有限或非法类型 / non finite or an illegal type
    FC_DL_RtdLinearization := FALSE; // 函数返回失败 / the function returns failure
    RETURN; // 早退 / early return
END_IF

// 段 2｜引线补偿与阻值域闸 / segment 2, lead compensation and the resistance domain gate
_fRUse := fROhm - fLeadOhm; // 扣除引线电阻 / subtract the lead resistance
IF (_fRUse < _fRMin) OR (_fRUse > _fRMax) THEN // 阻值越出测温域 / the resistance is outside the domain
    bOutOfRange := TRUE; // 置越域标志 / raise the out of range flag
    fTempC := 0.0; // 出口取安全侧零（R127）/ the outlet takes the safe side zero
    FC_DL_RtdLinearization := TRUE; // 函数返回成功（越域但可观测）/ the function returns success
    RETURN; // 早退 / early return
END_IF
IF _fRUse <= 0.0 THEN // 有效阻值非正（被引线补偿过度扣除，防御性保留）/ the effective resistance is void, kept as a defence
    bInvalid := TRUE; // 置无效标志 / raise the invalid flag
    FC_DL_RtdLinearization := FALSE; // 函数返回失败 / the function returns failure
    RETURN; // 早退 / early return
END_IF
_fRel := _fRUse / _fR0; // 相对阻值，除子为标称阻值常量已证非零 / the relative resistance, the divisor is the proven constant

// 段 3｜正温段二次方程求根 / segment 3, the positive branch quadratic root
_fDisc := _fA * _fA - 4.0 * _fB * (1.0 - _fRel); // 判别式 A^2 - 4B(1-r) / the discriminant
IF _fDisc < 0.0 THEN // 判别式为负，方程无实根 / a negative discriminant has no real root
    bInvalid := TRUE; // 置无效标志 / raise the invalid flag
    FC_DL_RtdLinearization := FALSE; // 函数返回失败 / the function returns failure
    RETURN; // 早退 / early return
END_IF
_fTPos := (-_fA + SQRT(_fDisc)) / (2.0 * _fB); // 求根公式取正根支，除子 2B 为负常量已证非零 / the root, the divisor is the proven negative constant
IF _fTPos >= 0.0 THEN // 正温段命中 / the positive branch hit
    fTempC := _fTPos; // 出口取正温根 / the outlet takes the positive root
    FC_DL_RtdLinearization := TRUE; // 函数返回成功 / the function returns success
    RETURN; // 早退 / early return
END_IF

// 段 4｜负温段定点迭代：T = (r - 1 - B·T^2 - C·(T-100)·T^3) / A（幂次显式乘法展开）/ segment 4, the negative branch fixed point iteration with explicit multiplications
_fTIt := -100.0; // 迭代初值取域中点 / the iterate starts at the domain mid point
_bConv := FALSE; // 收敛标志预置假 / preset the convergence flag to false
_nI := 0; // 守护游标清零 / clear the guard cursor
WHILE (_nI < 60) AND (NOT _bConv) DO // 双重守护：次数上限与收敛判据 / the dual guard on the count and the convergence
    _nI := _nI + 1; // 守护游标递增 / increment the guard
    _fTNext := (_fRel - 1.0 - _fB * _fTIt * _fTIt - _fC * (_fTIt - 100.0) * _fTIt * _fTIt * _fTIt) / _fA; // 定点迭代式，除子 A 为正常量已证非零 / the iteration step, the divisor is the proven positive constant
    _fDlt := ABS(_fTNext - _fTIt); // 步差 / the step difference
    _fTIt := _fTNext; // 推进迭代值 / advance the iterate
    IF _fDlt < 1.0E-9 THEN // 收敛达标 / the convergence is reached
        _bConv := TRUE; // 置收敛标志 / raise the convergence flag
    END_IF
END_WHILE
IF (NOT _bConv) OR (_fTIt < -200.0) OR (_fTIt >= 0.0) THEN // 不收敛或迭代跑出负温域 / no convergence or the iterate left the negative domain
    bInvalid := TRUE; // 置无效标志 / raise the invalid flag
    FC_DL_RtdLinearization := FALSE; // 函数返回失败 / the function returns failure
    RETURN; // 早退 / early return
END_IF
fTempC := _fTIt; // 出口取负温收敛值 / the outlet takes the converged negative value
FC_DL_RtdLinearization := TRUE; // 函数返回成功 / the function returns success
END_FUNCTION

(* ---- FC_DL_RunningSumCalc.st ---- *)
(*
  ==================================================================
  组件名 Component  : FC_DL_RunningSumCalc
  分类   Category   : DL_MathData
  前缀   Naming     : FC_DL_ ｜ b/n/u/f/t/e/st 类型前缀制（R265）
  码位   Code ID    : 16#0001_0668（故障级）｜ 16#0001_0669（信息级）
  版本   Version    : 1.0.0
  复杂度 Complexity  : 中
  功能   Purpose    : LREAL 运行累加和：Kahan 补偿求和防长序列累积误差，非
                      有限闸冻结状态，DINT 拍数饱和计数；供产期能耗累计、
                      批次总量计量、运行时长折算等调用方使用。
  开源溯源 Origin    : T0 统计族补口（内部来源，零检索）；Kahan 补偿求和为
                      公共领域算法（Kahan 1965）；增量式运行口径 + 非有限闸
                      为本库扩展，零代码复制。
  许可证 License    : MIT
  参考   Reference  : IEC 61131-3:2013 §6.6 算术运算符；Kahan 补偿求和
                      （Kahan 1965，公共领域算法）
  平台   Platform   : 纯 IEC 61131-3（四则 / 比较），三平台通用
  依赖   Depends    : 无（零委托、零库件）
  分工声明 Split     : FC_DL_SignalStatistics（窗口统计族，批内全量重算）为
                      互补件（互引）；本件为逐拍增量式运行口径（状态外置
                      结构体），统计族为窗内批处理口径，职责不同（R216）。
  归属 Ownership     : ST_DL_RunningSumState 属主为本文件（全库唯一定义，
                      R264）；引用件只引用不重声明。状态经 VAR_IN_OUT 外置，
                      本件零内部记忆量（FC 无实例态，纯 IEC 口径）。
  ------------------------------------------------------------------
  边界 Boundary     :
                      一 状态外置契约：累计状态（主和 / 补偿项 / 拍数）由
                         调用方持有（ST_DL_RunningSumState 实例经 VAR_IN_OUT
                         传入），本件零内部记忆量；调用方须每拍以同一实例
                         调用，跨实例混用即口径破坏（头注释声明，不做运行
                         期甄别——FC 无法取得实例身份，无永假防御）；
                      二 非有限闸：fSample 非有限（NaN / ±Inf）→ 故障级
                         0668 + 状态冻结（主和 / 补偿 / 拍数本拍不动）+
                         bValid = FALSE + bError = TRUE；nMaxScans < 1
                         （组态非法）出口组合同形（本拍不累加、状态不动、
                         三件套），合并一码（反证句见码表）；
                      三 Kahan 补偿链：y = fSample − fComp；t = fSum + y；
                         fComp = (t − fSum) − y；fSum = t（防长序列累积
                         误差，每拍补偿项回吸）；
                      四 结果复检：Kahan 后 fSum 非有限（理论上不可达的
                         兜底，R258）→ 同码 0668 + 状态冻结 + 三件套；
                      五 拍数饱和（信息级 0669）：nScans 已达 nMaxScans 后
                         拍数计数饱和钳位不再推进，累加本身继续（拍数是
                         审计量不是累加门槛），置信息级 0669 不置 bError；
                      六 bReset 电平复位：主和 / 补偿 / 拍数 / 冻结标记
                         全量清账（复位优先于累加，回夹路径显式清账）；
                      七 无定时器、无边沿实例；无除法；无全局、无外部
                         变量、无物理地址。
  错误码 Codes      :
    16#0001_0668【故障级】fSample 非有限（状态冻结）或 nMaxScans < 1（组态
                         非法）或结果复检命中非有限（三场景出口同形，合并一码）
    16#0001_0669【信息级】拍数已达 nMaxScans 饱和钳位（累加继续，不置 bError）
  码位反证 Note     :
    0668 合并三场景（样本非有限 / 拍数上限组态非法 / 结果复检命中）的理由：
    三场景出口组合完全相同（状态四元组本拍不动、bValid = FALSE、bError =
    TRUE），三组以内输出无法唯一还原该场景，按 R90 不另立码；0669 与 0668
    分立：0669 出口 bValid = TRUE（累加继续），bValid 可唯一区分。
  验收 Acceptance   :
    算法已证（脚本）：未跑 ｜ 编译器已证（三平台）：未跑
    V1 累加 1.0 × 10 拍 → fSum = 10.0、nScans = 10
    V2 长序列误差向量：1.0E16 起 +1.0 累加 1000 拍 → Kahan fSum 精度优于
       朴素累加（与 FC_DL_SignalStatistics 直和对比断言）
    V3 fSample = NaN 单拍 → 码 0668 + fSum 不动 + bError = TRUE，下一拍
       恢复正常样本继续累加（NaN 输入冻结不粘滞）
    V4 nMaxScans = 5、累加 8 拍 → nScans = 5（饱和）、fSum 照常推进、
       码 0669（bError = FALSE）
    V5 nMaxScans = 0 → 码 0668 + 状态不动
    V6 bReset 一拍 → fSum / fComp / nScans 全量清零
  修订记录 Revision  :
    2026-11-21  v1.0.0  R64 首版（批 2 · 序号 7，T0 统计族补口，Kahan 增量口径）
  ==================================================================
*)
TYPE ST_DL_RunningSumState :
STRUCT
    fSum   : LREAL := 0.0; // Kahan 主和 [工程单位] / the kahan main sum
    fComp  : LREAL := 0.0; // Kahan 补偿项 [工程单位]（每拍回吸损失）/ the kahan compensation term
    nScans : DINT   := 0;  // 累计拍数 [拍]（饱和上限 nMaxScans）/ the accumulated scan count saturated at the ceiling
    bFrozen: BOOL   := FALSE; // 状态冻结标记（非有限冻结期累计挂起）/ the frozen flag suspending the accumulation
END_STRUCT
END_TYPE

FUNCTION FC_DL_RunningSumCalc : BOOL
VAR_IN_OUT
    stState : ST_DL_RunningSumState; // 累计状态（调用方持有，须每拍同一实例）/ the accumulation state owned by the caller with the same instance every scan
END_VAR
VAR_INPUT
    fSample   : LREAL := 0.0; // 本拍样本 [工程单位]，必须有限 / the sample of this scan, must be finite
    nMaxScans : DINT   := 0;  // 拍数饱和上限 [拍]，须 ≥ 1，0 = 未组态（判故障）/ the scan ceiling, at least one, zero means unconfigured
    bReset    : BOOL  := FALSE; // 复位电平，TRUE 拍全量清账（复位优先于累加）/ the reset level clearing the whole state first
END_VAR
VAR_OUTPUT
    fSum   : LREAL; // 累加和出口 [工程单位] / the running sum outlet
    nScans : DINT;  // 累计拍数出口 [拍]（饱和口径）/ the scan count outlet saturated
    bValid : BOOL;  // 结果可用 [-] / the result usable flag
    eErr   : UDINT; // 错误码，0 = 正常 / the error code, zero is ok
    bError : BOOL;  // 故障标志（故障级码同拍置位，R45 配对）/ the fault flag raised with a fault level code
END_VAR
VAR
    fY : LREAL := 0.0; // Kahan 增量工作副本（样本 − 补偿）[工程单位] / the kahan increment copy of the sample minus the compensation
    fT : LREAL := 0.0; // Kahan 中间和工作副本 [工程单位] / the kahan intermediate sum copy
END_VAR  // R64 结构补齐：VAR 段缺失的 END_VAR（门禁机械修复）
VAR CONSTANT
    DL_RSC_ZERO : LREAL := 0.0; // 实数零常量 [工程单位] / the real zero constant
    DL_RSC_ZEROI: DINT   := 0;  // 整型零常量 [拍] / the integer zero constant
    DL_RSC_ONEI : DINT   := 1;  // 整型一常量 [拍] / the integer one constant
END_VAR

// 段 1｜返回值与全部出口预置安全值（R45 四段式第一段）/ segment 1, the preset of the return and all outlets
FC_DL_RunningSumCalc := FALSE; // 返回值预置假 / preset the return false
fSum := stState.fSum; // 和出口预置为现行状态值（冻结 / 复位口径的基线）[工程单位] / preset the sum outlet from the current state
nScans := stState.nScans; // 拍数出口预置为现行状态值 [拍] / preset the count outlet from the current state
bValid := FALSE; // 可用标志预置假 / preset the validity false
eErr := 16#0000_0000; // 错误码预置正常 / preset the code to ok
bError := FALSE; // 故障标志预置假 / preset the fault flag false
fY := DL_RSC_ZERO; // Kahan 增量预置零 [工程单位] / preset the kahan increment zero
fT := DL_RSC_ZERO; // Kahan 中间和预置零 [工程单位] / preset the kahan intermediate zero

// 段 2｜复位优先段（边界六：全量清账，复位优先于累加与一切闸）/ segment 2, the reset first with the full clearing
IF bReset THEN // 复位电平有效 / the reset level is active
    stState.fSum := DL_RSC_ZERO; // 主和清账 [工程单位] / clear the main sum
    stState.fComp := DL_RSC_ZERO; // 补偿项清账 [工程单位] / clear the compensation
    stState.nScans := DL_RSC_ZEROI; // 拍数清账 [拍] / clear the scan count
    stState.bFrozen := FALSE; // 冻结标记清账 / clear the frozen flag
    fSum := DL_RSC_ZERO; // 和出口同步清零 [工程单位] / sync the sum outlet zero
    nScans := DL_RSC_ZEROI; // 拍数出口同步清零 [拍] / sync the count outlet zero
    bValid := TRUE; // 复位是合法可用结果 / the reset is a legit usable result
    FC_DL_RunningSumCalc := TRUE; // 返回成功 / return success
    RETURN; // 早退（复位拍不累加）/ early return, no accumulation on the reset scan
END_IF

// 段 3｜非有限闸与组态闸（边界二：两场景出口同形合并一码，状态冻结）/ segment 3, the finiteness gate and the configuration gate freezing the state
IF (fSample <> fSample) OR ((fSample - fSample) <> (fSample - fSample))
OR (nMaxScans < DL_RSC_ONEI) THEN // 样本非有限或拍数上限组态非法 / the sample is not finite or the ceiling is misconfigured
    stState.bFrozen := TRUE; // 置状态冻结（本拍累计挂起）/ raise the frozen flag
    eErr := 16#0001_0668; // 故障级：非有限或组态非法（合并一码，R90）/ fault grade under the merged code
    bError := TRUE; // 同拍置故障标志（R45 配对）/ raise the fault flag on the same scan
    bValid := FALSE; // 结果不可用 / the result is not usable
    RETURN; // 早退，状态四元组本拍不动 / early return, the state untouched this scan
END_IF

// 段 4｜Kahan 补偿累加（边界三；冻结期挂起，恢复后自动续计）/ segment 4, the kahan compensated accumulation
IF NOT stState.bFrozen THEN // 未冻结才累加 / accumulate only when not frozen
    fY := fSample - stState.fComp; // 增量 = 样本 − 补偿项 [工程单位] / the increment of the sample minus the compensation
    fT := stState.fSum + fY; // 中间和 [工程单位] / the intermediate sum
    stState.fComp := (fT - stState.fSum) - fY; // 补偿项回吸本轮舍入损失 [工程单位] / the compensation sucking back the rounding loss
    stState.fSum := fT; // 主和推进 [工程单位] / advance the main sum
    IF stState.nScans < nMaxScans THEN // 拍数未达上限 / the count below the ceiling
        stState.nScans := stState.nScans + DL_RSC_ONEI; // 拍数推进 [拍] / advance the scan count
    ELSE // 拍数已达上限：饱和钳位 + 信息级（累加继续，边界五）/ the count saturated with the info code, the accumulation continues
        eErr := 16#0001_0669; // 信息级：拍数饱和钳位（R285）/ informational, the count is saturated
        bError := FALSE; // 信息级不置故障标志 / keep the fault flag false, this is informational
    END_IF
ELSE // 冻结期（上拍非有限命中后本拍已过闸，自动解冻续计）/ the frozen period auto releases after the gate passed
    stState.bFrozen := FALSE; // 解冻（非有限输入冻结不粘滞，恢复路径可达）/ release the frozen flag, the recovery is reachable
    fY := fSample - stState.fComp; // 解冻拍照常累加 [工程单位] / accumulate as usual on the release scan
    fT := stState.fSum + fY; // 中间和 [工程单位] / the intermediate sum
    stState.fComp := (fT - stState.fSum) - fY; // 补偿项回吸 [工程单位] / the compensation
    stState.fSum := fT; // 主和推进 [工程单位] / advance the main sum
    IF stState.nScans < nMaxScans THEN // 拍数未达上限 / the count below the ceiling
        stState.nScans := stState.nScans + DL_RSC_ONEI; // 拍数推进 [拍] / advance the scan count
    ELSE // 拍数饱和（信息级，累加继续）/ the count saturated, the accumulation continues
        eErr := 16#0001_0669; // 信息级：拍数饱和钳位 / informational, the count is saturated
        bError := FALSE; // 信息级不置故障标志 / keep the fault flag false
    END_IF
END_IF

// 段 5｜结果复检兜底（边界四：理论上不可达，R258 三件套 + 状态冻结）/ segment 5, the result recheck with the three part fallback
IF (stState.fSum <> stState.fSum) OR ((stState.fSum - stState.fSum) <> (stState.fSum - stState.fSum)) THEN // 主和非有限（兜底防御）/ the main sum is not finite
    stState.bFrozen := TRUE; // 置状态冻结 / raise the frozen flag
    eErr := 16#0001_0668; // 故障级：结果复检命中（同形合并一码，R90）/ fault grade under the merged code
    bError := TRUE; // 置故障标志（R45 配对）/ raise the fault flag
    bValid := FALSE; // 结果不可用 / the result is not usable
    RETURN; // 早退，状态冻结 / early return with the state frozen
END_IF

// 段 6｜统一出口 / segment 6, the unified outlet
fSum := stState.fSum; // 和出口 [工程单位] / the sum outlet
nScans := stState.nScans; // 拍数出口 [拍] / the count outlet
bValid := TRUE; // 结果可用 / the result is usable
FC_DL_RunningSumCalc := TRUE; // 返回成功 / return success
END_FUNCTION
